// ST-FIX F23: wait until the RC left the state INITIALIZED of the previous enable
IF ( _restartReset )
THEN
  IF ( AxesGroup.Cyclic.RobToPlc.TelegramState <> TelegramState.INITIALIZED )
  THEN
    _restartReset := FALSE;
  END_IF
ELSE
CASE AxesGroup.Cyclic.RobToPlc.TelegramState  OF

         TelegramState.UNDEFINED : ;
         
         TelegramState.ERROR_161_TELEGRAM_CONTROL_MISMATCH_TELEGRAM_STATE..TelegramState.ERROR_172_TELEGRAM_NUMBER_NOT_SUPPORTED:

           // ST-FIX F79: remember the error state for the init timeout
           _initErrorState := AxesGroup.Cyclic.RobToPlc.TelegramState;

           // clear error
           AxesGroup.Cyclic.PlcToRob.Control := ControlHalfByte.ACK_ERROR;        
           AxesGroup.Cyclic.PlcToRob.Control := ControlHalfByte.RESET; // always a reset, so that on the robot side the ACR is reseted         

         TelegramState.ERROR_173_SERVER_CONNECTION_LOST:

           // Reset interface including the ACR register on server side
           AxesGroup.Cyclic.PlcToRob.Control := ControlHalfByte.RESET;        
           
         TelegramState.READY_TO_RESUME :  
         
           // Resume
           AxesGroup.Cyclic.PlcToRob.Control := ControlHalfByte.RESUME;        
         
         TelegramState.READY_FOR_INITIALIZATION: 

           // Request initialization
           AxesGroup.Cyclic.PlcToRob.Control := ControlHalfByte.INITIALIZE;
           
         TelegramState.INITIALIZED: 

           // Reset Telegram Control 
           AxesGroup.Cyclic.PlcToRob.Control := ControlHalfByte.NONE;
           
           // Check SRCI Version is compatible ? 
           IF ( AxesGroup.Cyclic.RobToPlc.SRCIVersion.MajorVersion = RobotLibraryConstants.SRCIVersion.MajorVersion )
           THEN
             // set timeout
             SetTimeout(PT := _timeoutCmd, rTimer := _timerCmd);
             // inc step counter
            _stepCmd := _stepCmd + 1; 
           ELSE
             // set error 
             ErrorID     := RobotLibraryErrorIdEnum.ERR_SRCI_MAJOR_VERSION_INCOMPATIBLE_0x80A4;
             ErrorAddTxt := CONCAT('_stepCmd = ' , DINT_TO_STRING(_stepCmd));
           END_IF

       ELSE
         // TelegrammState in error          
         SetError( ErrorID := RobotLibraryErrorIdEnum.ERR_INIT_LOST_UNKNOWN_0x80A2, Overwrite := TRUE ); // ST-FIX F65: unknown state (16#A2 is the RI error of the RC)
           // Create log entry
           CreateLogMessagePara1 ( Timestamp   := SystemTime,
                                   MessageType := MessageType.CMD,
                                   Severity    := Severity.ERROR,
                                   MessageCode := ErrorID,
                                   MessageText := 'Initialization lost: unknown telegram state {1}',
                                   Para1       := TELEGRAM_STATE_TO_STRING(AxesGroup.Cyclic.RobToPlc.TelegramState));
         ErrorAddTxt := CONCAT('_stepCmd = ' , DINT_TO_STRING(_stepCmd));
       END_CASE
END_IF

       // timeout exceeded ? 
       IF (CheckTimeout(_timerCmd) = RobotLibraryConstants.OK)
       THEN
         // Check Telegram State error ? 
         IF (( AxesGroup.Cyclic.RobToPlc.TelegramState >= TelegramState.ERROR_161_TELEGRAM_CONTROL_MISMATCH_TELEGRAM_STATE ) AND // ST-FIX F15
             ( AxesGroup.Cyclic.RobToPlc.TelegramState <= TelegramState.ERROR_173_SERVER_CONNECTION_LOST                   ))
         THEN
           ErrorID     := AxesGroup.Cyclic.RobToPlc.TelegramState;
           ErrorAddTxt := CONCAT('_stepCmd = ' , DINT_TO_STRING(_stepCmd));
         ELSIF ( _initErrorState <> TelegramState.UNDEFINED ) // ST-FIX F79: error state seen during the initialization
         THEN
           ErrorID     := _initErrorState;
           ErrorAddTxt := CONCAT('_stepCmd = ' , DINT_TO_STRING(_stepCmd));
         ELSE
           ErrorID     := RobotLibraryErrorIdEnum.ERR_TIMEOUT_CMD;
           ErrorAddTxt := CONCAT('_stepCmd = ' , DINT_TO_STRING(_stepCmd));
         END_IF
       END_IF

       
  02: IF (( NOT _readMessages.Busy  ) AND 
          ( NOT _readMessages.Error )) 
      THEN
        // start function block
       _readMessages.Enable := TRUE;
       _readMessages.ParCmd.MsgID := 0;
       _readMessages.ParCmd.MessageLevel := _parCfg.Rob.Parameter.MessageLevel;
        
        // set timeout
        SetTimeout(PT := _timeoutCmd, rTimer := _timerCmd);
        // inc step counter
       _stepCmd := _stepCmd + 1;       
      ELSE
        // check error ? 
        IF (_readMessages.Error)
        THEN
          ErrorID     := _readMessages.ErrorID;
          ErrorAddTxt := _readMessages.ErrorAddTxt;;
        END_IF  
        // timeout exceeded ? 
        IF (CheckTimeout(_timerCmd) = RobotLibraryConstants.OK)
        THEN
          ErrorID     := RobotLibraryErrorIdEnum.ERR_TIMEOUT_CMD;
          ErrorAddTxt := CONCAT('_stepCmd = ' , DINT_TO_STRING(_stepCmd));
        END_IF
      END_IF
  
  03: IF ((     _readMessages.Enabled ) AND
          ( NOT _readMessages.Error   ))
      THEN       
        // --------------------------------------------------------------- 
        // !!! ReadMessages must stay active for the Message mechanism !!!
        // --------------------------------------------------------------- 
        // ReadMessages.Enable := FALSE;  
        // set timeout
        SetTimeout(PT := _timeoutCmd, rTimer := _timerCmd);
        // inc step counter
       _stepCmd := _stepCmd + 1;
      ELSE
         // check error ? 
         IF (_readMessages.Error)
         THEN
           ErrorID     := _readMessages.ErrorID;
           ErrorAddTxt := _readMessages.ErrorAddTxt;;
         END_IF  
       
         // timeout exceeded ? 
         IF (CheckTimeout(_timerCmd) = RobotLibraryConstants.OK)
         THEN
           ErrorID     := RobotLibraryErrorIdEnum.ERR_TIMEOUT_CMD;
           ErrorAddTxt := CONCAT('_stepCmd = ' , DINT_TO_STRING(_stepCmd));
         END_IF
       END_IF       
       
       
  04: IF (( NOT _exchangeConfiguration.Busy  ) AND 
          ( NOT _exchangeConfiguration.Error ))
      THEN
        // set command parameter
       _exchangeConfiguration.ParCmd.LogLevel                           :=  LogLevel; 
       _exchangeConfiguration.ParCmd.WaitAtBlendingZone                 := _parCfg.Rob.Parameter.WaitAtBlendingZone;
       _exchangeConfiguration.ParCmd.AllowSecSeqWhileSubprogram         := _parCfg.Rob.Parameter.AllowSecSeqWhileSubprogram;
       _exchangeConfiguration.ParCmd.AllowDynamicBlending               := _parCfg.Rob.Parameter.AllowDynamicBlending;
       _exchangeConfiguration.ParCmd.DelayTime                          := _parCfg.Rob.Parameter.DelayTime;
       _exchangeConfiguration.ParCmd.WaitForNrOfCmd                     := _parCfg.Rob.Parameter.WaitForNrOfCmd;
       _exchangeConfiguration.ParCmd.LifeSignTimeOut                    :=  TIME_TO_UINT(_parCfg.Com.LifeSignTimeOut);
       _exchangeConfiguration.ParCmd.SyncDelay                          := _parCfg.Rob.Parameter.SyncDelay;
       _exchangeConfiguration.ParCmd.SyncReaction                       := _parCfg.Rob.Parameter.SyncReaction;
       _exchangeConfiguration.ParCmd.DataEnableSync                     :=  SyncModesToDataEnableSync(Value := _parCfg.Plc.Parameter.SynchronizationModes);
       _exchangeConfiguration.ParCmd.DataInSync.ToolsInSync             :=  FALSE;
       _exchangeConfiguration.ParCmd.DataInSync.FramesInSync            :=  FALSE;
       _exchangeConfiguration.ParCmd.DataInSync.LoadsInSync             :=  FALSE;
       _exchangeConfiguration.ParCmd.DataInSync.WorkAreasInSync         :=  FALSE;
       _exchangeConfiguration.ParCmd.DataInSync.SoftwareLimitsInSync    :=  FALSE;
       _exchangeConfiguration.ParCmd.DataInSync.DefaultDynamicsInSync   :=  FALSE;
       _exchangeConfiguration.ParCmd.DataInSync.ReferenceDynamicsInSync :=  FALSE;         
       
        // start function block
       _exchangeConfiguration.Enable := TRUE;
        // set timeout
        SetTimeout(PT := _timeoutCmd, rTimer := _timerCmd);
        // inc step counter
       _stepCmd := _stepCmd + 1;       
      ELSE
        // check error ? 
        IF (_exchangeConfiguration.Error)
        THEN
          ErrorID     := _exchangeConfiguration.ErrorID;
          ErrorAddTxt := _exchangeConfiguration.ErrorAddTxt;;
        END_IF  
       
        // timeout exceeded ? 
        IF (CheckTimeout(_timerCmd) = RobotLibraryConstants.OK)
        THEN
          ErrorID     := RobotLibraryErrorIdEnum.ERR_TIMEOUT_CMD;
          ErrorAddTxt := CONCAT('_stepCmd = ' , DINT_TO_STRING(_stepCmd));
        END_IF
      END_IF
  
  
  05: IF ((     _exchangeConfiguration.Enabled ) AND
          ( NOT _exchangeConfiguration.Error   ))
      THEN     
        // --------------------------------------------------------------------- 
        // !!! ExchangeConfiguration must stay active for the Sync mechanism !!!
        // --------------------------------------------------------------------- 
        // ExchangeConfiguration.Enable := FALSE;  
        // set timeout
        SetTimeout(PT := _timeoutCmd, rTimer := _timerCmd);
        // inc step counter
       _stepCmd := _stepCmd + 1;       
      ELSE
        // check error ? 
        IF (_exchangeConfiguration.Error)
        THEN
          ErrorID     := _exchangeConfiguration.ErrorID;
          ErrorAddTxt := _exchangeConfiguration.ErrorAddTxt;;
        END_IF  
       
        // timeout exceeded ? 
        IF (CheckTimeout(_timerCmd) = RobotLibraryConstants.OK)
        THEN
          ErrorID     := RobotLibraryErrorIdEnum.ERR_TIMEOUT_CMD;
          ErrorAddTxt := CONCAT('_stepCmd = ' , DINT_TO_STRING(_stepCmd));
        END_IF
      END_IF

       
  06: IF (( NOT _readRobotData.Busy  ) AND 
          ( NOT _readRobotData.Error )) 
      THEN
        // start function block
       _readRobotData.Execute := TRUE;
        // set timeout
        SetTimeout(PT := _timeoutCmd, rTimer := _timerCmd);
        // inc step counter
       _stepCmd := _stepCmd + 1;       
      ELSE
        // check error ? 
        IF (_readRobotData.Error)
        THEN
          ErrorID     := _readRobotData.ErrorID;
          ErrorAddTxt := _readRobotData.ErrorAddTxt;;
        END_IF  
        // timeout exceeded ? 
        IF (CheckTimeout(_timerCmd) = RobotLibraryConstants.OK)
        THEN
          ErrorID     := RobotLibraryErrorIdEnum.ERR_TIMEOUT_CMD;
          ErrorAddTxt := CONCAT('_stepCmd = ' , DINT_TO_STRING(_stepCmd));
        END_IF
      END_IF
    
  
  07: IF ((     _readRobotData.Done  ) AND
          ( NOT _readRobotData.Busy  ) AND
          ( NOT _readRobotData.Error ))          
      THEN       
        // set initialized flag
        Initialized := TRUE;       
        // start function block
       _readRobotData.Execute := FALSE;
        // set timeout
        SetTimeout(PT := _timeoutCmd, rTimer := _timerCmd);
        // inc step counter
       _stepCmd := _stepCmd + 1;
       ELSE
         // check error ? 
         IF (_readRobotData.Error)
         THEN
           ErrorID     := _readRobotData.ErrorID;
           ErrorAddTxt := _readRobotData.ErrorAddTxt;;
         END_IF  
       
         // timeout exceeded ? 
         IF (CheckTimeout(_timerCmd) = RobotLibraryConstants.OK)
         THEN
           ErrorID     := RobotLibraryErrorIdEnum.ERR_TIMEOUT_CMD;
           ErrorAddTxt := CONCAT('_stepCmd = ' , DINT_TO_STRING(_stepCmd));
         END_IF
       END_IF

       
  08:  // Update Initialized state
       // ST-FIX F131: Initialized stays TRUE while Synchronized (RI state "Synchronized" includes the
       // initialization); otherwise CheckParameterChanged did not run while synchronized
       Initialized := NOT Error;
       // ST-FIX F29: the next line overwrote the error check above
       // Initialized := NOT Synchronized;

       // Wait for task disable
       IF ( NOT Enable)
       THEN
         // Reset active command register
         AxesGroup.Acyclic.ActiveCommandRegister.Reset();
         // reset internal variables
         Reset(AxesGroup := AxesGroup);
         // Reset step counter
        _stepCmd := 0;         
         // finished okay
         OnExecRun := RobotLibraryConstants.OK;
       END_IF  

       
ELSE
  // invalid step
  ErrorID     := RobotLibraryErrorIdEnum.ERR_INVALID_STEP;
  ErrorAddTxt := CONCAT('_stepCmd = ' , DINT_TO_STRING(_stepCmd));
END_CASE
END_METHOD

METHOD PROTECTED ParseRecvPayload
VAR_IN_OUT
  /// Robot assignment of function
  AxesGroup   : AxesGroup;
  /// Inputs of PLC for communication from RC
  RobotInData : ARRAY[*] OF BYTE;
END_VAR
// reset all variables and payload
RecvData.Reset();
// Call RecvData FB, update payload and size 
RecvData(Payload := RobotInData, PayloadSize := ROBOT_IN_DATA_SIZE);

// check new data to receive ? 
// ST-FIX F140: also new data of the 2nd sequence
IF ( Telegram.RobToPlc.Sequence[0].Header.SEQ_ACK <> AxesGroup.State.LastACK[0] ) OR
   ( Telegram.RobToPlc.Sequence[1].Header.SEQ_ACK <> AxesGroup.State.LastACK[1] )
THEN
  // delete old telegram data 
  SysDepMemSet(pDest := ADR(Telegram.RobToPlc), Value := 0 , DataLen := SIZEOF(Telegram.RobToPlc));
END_IF


ParseRecvPayloadHeader        ( AxesGroup := AxesGroup);
ParseRecvPayloadCyclic        ( AxesGroup := AxesGroup);
ParseRecvPayloadCyclicOptional( AxesGroup := AxesGroup);
ParseRecvPayloadSequence      ( AxesGroup := AxesGroup);
ParseRecvPayloadFooter        ( AxesGroup := AxesGroup);
ParseRecvPayloadLogging       ( AxesGroup := AxesGroup);


AxesGroup.State.LastACK[0] := Telegram.RobToPlc.Sequence[0].Header.SEQ_ACK; 
AxesGroup.State.LastACK[1] := Telegram.RobToPlc.Sequence[1].Header.SEQ_ACK;
END_METHOD

METHOD PROTECTED ParseRecvPayloadCyclic
VAR_IN_OUT
  /// Robot assignment of function
  AxesGroup: AxesGroup;
END_VAR
END_METHOD

METHOD PROTECTED ParseRecvPayloadCyclicOptional
VAR_IN_OUT
  /// Robot assignment of function
  AxesGroup    : AxesGroup;
END_VAR

VAR 
  /// internal index for loops
 _idx : DINT;
END_VAR
// AxesGroup.OptionalCyclic.RobToPlc.SubProgramData {{{
IF ( AxesGroup.CyclicOptional.RobToPlc.SubProgramData.Active )
THEN
  FOR _idx := 0 TO  RobotLibraryConstants.CYCLIC_SUB_PROGRAM_DATA_MAX (* ST-FIX F179 *)
  DO
    Telegram.RobToPlc.CyclicOptional.SubProgramData.Data[_idx] := RecvData.GetByte(); 
  END_FOR
END_IF
// }}}
  
// AxesGroup.OptionalCyclic.RobToPlc.CartesianPos {{{
IF ( AxesGroup.CyclicOptional.RobToPlc.CartesianPosition.Active )
THEN
  Telegram.RobToPlc.CyclicOptional.CartesianPosition.X                    := RecvData.GetReal();
  Telegram.RobToPlc.CyclicOptional.CartesianPosition.Y                    := RecvData.GetReal();
  Telegram.RobToPlc.CyclicOptional.CartesianPosition.Z                    := RecvData.GetReal();
  Telegram.RobToPlc.CyclicOptional.CartesianPosition.Rx                   := RecvData.GetReal();
  Telegram.RobToPlc.CyclicOptional.CartesianPosition.Ry                   := RecvData.GetReal();
  Telegram.RobToPlc.CyclicOptional.CartesianPosition.Rz                   := RecvData.GetReal();
  Telegram.RobToPlc.CyclicOptional.CartesianPosition.Config               := RecvData.GetWord();
  Telegram.RobToPlc.CyclicOptional.CartesianPosition.Turns_J2_J1          := RecvData.GetByte();
  Telegram.RobToPlc.CyclicOptional.CartesianPosition.Turns_J4_J3          := RecvData.GetByte();
  Telegram.RobToPlc.CyclicOptional.CartesianPosition.Turns_J6_J5          := RecvData.GetByte();
  Telegram.RobToPlc.CyclicOptional.CartesianPosition.Turns_E1             := RecvData.GetByte();  
  Telegram.RobToPlc.CyclicOptional.CartesianPosition.E1                   := RecvData.GetReal();  
  Telegram.RobToPlc.CyclicOptional.CartesianPosition.ToolNo               := RecvData.GetUsint();
  Telegram.RobToPlc.CyclicOptional.CartesianPosition.FrameNo              := RecvData.GetUsint();
  Telegram.RobToPlc.CyclicOptional.CartesianPosition.CurrentlyUsedToolNo  := RecvData.GetUsint();
  Telegram.RobToPlc.CyclicOptional.CartesianPosition.CurrentlyUsedFrameNo := RecvData.GetUsint();
  Telegram.RobToPlc.CyclicOptional.CartesianPosition.Reserve_1            := RecvData.GetByte();
  Telegram.RobToPlc.CyclicOptional.CartesianPosition.Reserve_2            := RecvData.GetByte();  
END_IF
// }}}

// AxesGroup.OptionalCyclic.RobToPlc.JointPosition {{{
IF ( AxesGroup.CyclicOptional.RobToPlc.JointPosition.Active )
THEN
  Telegram.RobToPlc.CyclicOptional.JointPosition.J1         := RecvData.GetReal();
  Telegram.RobToPlc.CyclicOptional.JointPosition.J2         := RecvData.GetReal();
  Telegram.RobToPlc.CyclicOptional.JointPosition.J3         := RecvData.GetReal();
  Telegram.RobToPlc.CyclicOptional.JointPosition.J4         := RecvData.GetReal();
  Telegram.RobToPlc.CyclicOptional.JointPosition.J5         := RecvData.GetReal();
  Telegram.RobToPlc.CyclicOptional.JointPosition.J6         := RecvData.GetReal();
  Telegram.RobToPlc.CyclicOptional.JointPosition.E1         := RecvData.GetReal();
  Telegram.RobToPlc.CyclicOptional.JointPosition.E1_Reserve := RecvData.GetWord();
END_IF  
// }}}

// AxesGroup.OptionalCyclic.RobToPlc.CartesianForce {{{
IF ( AxesGroup.CyclicOptional.RobToPlc.Force.Active )
THEN
  Telegram.RobToPlc.CyclicOptional.Force.X  := RecvData.GetReal();
  Telegram.RobToPlc.CyclicOptional.Force.Y  := RecvData.GetReal();
  Telegram.RobToPlc.CyclicOptional.Force.Z  := RecvData.GetReal();
  Telegram.RobToPlc.CyclicOptional.Force.Rx := RecvData.GetReal();
  Telegram.RobToPlc.CyclicOptional.Force.Ry := RecvData.GetReal();
  Telegram.RobToPlc.CyclicOptional.Force.Rz := RecvData.GetReal();
END_IF  
// }}}    
  
// AxesGroup.OptionalCyclic.RobToPlc.Current {{{
IF ( AxesGroup.CyclicOptional.RobToPlc.Current.Active )
THEN
  Telegram.RobToPlc.CyclicOptional.Current.J1  := RecvData.GetReal();
  Telegram.RobToPlc.CyclicOptional.Current.J2  := RecvData.GetReal();
  Telegram.RobToPlc.CyclicOptional.Current.J3  := RecvData.GetReal();
  Telegram.RobToPlc.CyclicOptional.Current.J4  := RecvData.GetReal();
  Telegram.RobToPlc.CyclicOptional.Current.J5  := RecvData.GetReal();
  Telegram.RobToPlc.CyclicOptional.Current.J6  := RecvData.GetReal();
END_IF    
  
// AxesGroup.OptionalCyclic.RobToPlc.CartesianPosExt {{{
IF ( AxesGroup.CyclicOptional.RobToPlc.CartesianPositionExt.Active )
THEN
  Telegram.RobToPlc.CyclicOptional.CartesianPositionExt.E2 := RecvData.GetReal();
  Telegram.RobToPlc.CyclicOptional.CartesianPositionExt.E3 := RecvData.GetReal();
  Telegram.RobToPlc.CyclicOptional.CartesianPositionExt.E4 := RecvData.GetReal();
  Telegram.RobToPlc.CyclicOptional.CartesianPositionExt.E5 := RecvData.GetReal();
  Telegram.RobToPlc.CyclicOptional.CartesianPositionExt.E6 := RecvData.GetReal();
END_IF  
// }}}       
  
// AxesGroup.OptionalCyclic.RobToPlc.JointPosition {{{
IF ( AxesGroup.CyclicOptional.RobToPlc.JointPositionExt.Active )
THEN
  Telegram.RobToPlc.CyclicOptional.JointPositionExt.E2 := RecvData.GetReal();
  Telegram.RobToPlc.CyclicOptional.JointPositionExt.E3 := RecvData.GetReal();
  Telegram.RobToPlc.CyclicOptional.JointPositionExt.E4 := RecvData.GetReal();
  Telegram.RobToPlc.CyclicOptional.JointPositionExt.E5 := RecvData.GetReal();
  Telegram.RobToPlc.CyclicOptional.JointPositionExt.E6 := RecvData.GetReal();  
END_IF  
// }}}    
      
// AxesGroup.OptionalCyclic.RobToPlc.CartesianForceExt {{{
IF ( AxesGroup.CyclicOptional.RobToPlc.ForceExt.Active )
THEN
  Telegram.RobToPlc.CyclicOptional.ForceExt.E1  := RecvData.GetReal();
  Telegram.RobToPlc.CyclicOptional.ForceExt.E2  := RecvData.GetReal();
  Telegram.RobToPlc.CyclicOptional.ForceExt.E3  := RecvData.GetReal();
  Telegram.RobToPlc.CyclicOptional.ForceExt.E4  := RecvData.GetReal();
  Telegram.RobToPlc.CyclicOptional.ForceExt.E5  := RecvData.GetReal();
  Telegram.RobToPlc.CyclicOptional.ForceExt.E6  := RecvData.GetReal();
END_IF
// }}}    
  
// AxesGroup.OptionalCyclic.RobToPlc.CurrentExt {{{
IF ( AxesGroup.CyclicOptional.RobToPlc.CurrentExt.Active )
THEN
  Telegram.RobToPlc.CyclicOptional.CurrentExt.E1  := RecvData.GetReal();
  Telegram.RobToPlc.CyclicOptional.CurrentExt.E2  := RecvData.GetReal();
  Telegram.RobToPlc.CyclicOptional.CurrentExt.E3  := RecvData.GetReal();
  Telegram.RobToPlc.CyclicOptional.CurrentExt.E4  := RecvData.GetReal();
  Telegram.RobToPlc.CyclicOptional.CurrentExt.E5  := RecvData.GetReal();
  Telegram.RobToPlc.CyclicOptional.CurrentExt.E6  := RecvData.GetReal();
END_IF
// }}}
END_METHOD

METHOD PRIVATE ParseRecvPayloadFooter
VAR_IN_OUT
  /// Robot assignment of function
  AxesGroup : AxesGroup;
END_VAR
Telegram.RobToPlc.Footer.LifeSign := RecvData.GetLifeSignFooter();
END_METHOD

METHOD PROTECTED ParseRecvPayloadHeader
VAR_IN_OUT
  /// Robot assignment of function
  AxesGroup    : AxesGroup;
END_VAR
// Version
Telegram.RobToPlc.Header.SRCIVersion := ByteToVersion(RecvData.GetByte());
// Connection alive signal
Telegram.RobToPlc.Header.LifeSign    := RecvData.GetHalfeByte2(IncPayloadPtr := TRUE);
// Reserved byte
Telegram.RobToPlc.Header.Reserved       := RecvData.GetByte();
// Initialization and Telegram control state
Telegram.RobToPlc.Header.TelegramState  := RecvData.GetUsint();
// Combination of various RA related states.
Telegram.RobToPlc.Header.StatusRobotArm := RecvData.GetDword();
// Actual override in percentage encoding 
Telegram.RobToPlc.Header.Override       := RecvData.GetUint();
END_METHOD

METHOD PRIVATE ParseRecvPayloadLogging
VAR_IN_OUT
  /// Robot assignment of function
  AxesGroup    : AxesGroup;
END_VAR

VAR
  /// internal sequence index for loops
  _seqIdx : DINT;
  /// internal fragment index for loops
  _fragIdx : DINT;
END_VAR
RETURN;
FOR _seqIdx := 0 TO AxesGroup.State.SequenceCountRecv
DO
  // check new data to receive ? 
  IF ( Telegram.RobToPlc.Sequence[_seqIdx].Header.SEQ_ACK <> AxesGroup.State.LastACK[_seqIdx]) 
  THEN
    // Check sequence payload > 0 ?    
    IF (Telegram.RobToPlc.Sequence[_seqIdx].Header.PayloadLength > 0)
    THEN
      // Create log entry
      CreateLogMessagePara4 ( Timestamp   := SystemTime,
                              MessageType := MessageType.CMD,
                              Severity    := Severity.DEBUG,
                              MessageCode := 0,
                              MessageText := 'RecvData: ACK = {1}, received Sequence [{2}] with PayloadLength = {3}, Lifesign = {4}',
                              Para1       :=  UINT_TO_STRING(Telegram.RobToPlc.Sequence[_seqIdx].Header.SEQ_ACK),
                              Para2       :=  DINT_TO_STRING(_seqIdx),
                              Para3       :=  UINT_TO_STRING(Telegram.RobToPlc.Sequence[_seqIdx].Header.PayloadLength),
                              Para4       :=  BYTE_TO_STRING(Telegram.RobToPlc.Header.LifeSign));
  
      FOR _fragIdx := 0 TO AxesGroup.State.FragmentCountRecv[_seqIdx] 
      DO
        // Check fragment payload > 0 ?    
        IF (Telegram.RobToPlc.Sequence[_seqIdx].Fragment[_fragIdx].Header.PayloadLength > 0)
        THEN
          // Create log entry
          CreateLogMessagePara5 ( Timestamp   := SystemTime,
                                  MessageType := MessageType.CMD,
                                  Severity    := Severity.DEBUG,
                                  MessageCode := 0,
                                  MessageText := 'RecvData: received Fragment [{1}] with PayloadLength = {2}, CmdID <{3}> , CmdState: {4}, Fragment-Action Bits: {5}',
                                  Para1       :=  DINT_TO_STRING(_fragIdx),
                                  Para2       :=  UINT_TO_STRING              (Telegram.RobToPlc.Sequence[_seqIdx].Fragment[_fragIdx].Header.PayloadLength),
                                  Para3       :=  DINT_TO_STRING              (Telegram.RobToPlc.Sequence[_seqIdx].Fragment[_fragIdx].Header.CmdID),
                                  Para4       :=  CMD_MESSAGE_STATE_TO_STRING (Telegram.RobToPlc.Sequence[_seqIdx].Fragment[_fragIdx].Command.Header.State),
                                  Para5       :=    FRAGMENT_ACTION_TO_STRING (Telegram.RobToPlc.Sequence[_seqIdx].Fragment[_fragIdx].Header.FragmentAction));
        END_IF
      END_FOR    
    END_IF
  END_IF
END_FOR
END_METHOD

METHOD PRIVATE ParseRecvPayloadSequence
VAR_IN_OUT
  /// Robot assignment of function
  AxesGroup        : AxesGroup;
END_VAR

VAR
  /// internal index
 _idx              : DINT;
  /// index for sequence
 _seqIdx           : DINT;
  /// index for fragment
 _fragIdx          : DINT; 
  /// current payload pointer for current fragment
 _payLoadPtr       : DINT;
  /// Amount of sequences
 _seqCount         : DINT;
  /// current payload pointer of the current sequence
 _seqPayloadPtr    : UINT; 
  /// ST-FIX F63: start of the payload of each sequence (behind its sequence header)
 _rcvStart         : ARRAY[0..1] OF DINT;
  /// ST-FIX F63: sequence that is processed first (lower Ack)
 _rcvFirst         : DINT;
  /// ST-FIX F63: loop counter over the sequences in Ack order
 _rcvOrderIdx      : DINT;
  /// ST-FIX F63: distance of the two Ack numbers
 _rcvDiff          : DINT;
END_VAR
// Check 2nd sequence active ? 
IF ( _parCfg.Com.TwoSequences )
THEN
 _seqCount := _seqCount + 1;
END_IF

// ST-FIX F63: read the headers of all sequences, each from its own address (Fig. 5-205)
FOR _seqIdx := 0 TO _seqCount
DO
  IF ( _seqIdx = PRIMARY_SEQUENCE )
  THEN
    RecvData.PayloadPtr := CalculateSequencePayloadStartAdr(AxesGroup := AxesGroup, 
                                                            Direction := ComDirection.ROB_TO_PLC,
                                                            Sequence  := SequenceFlag.PRIMARY_SEQUENCE);
  ELSE
    RecvData.PayloadPtr := CalculateSequencePayloadStartAdr(AxesGroup := AxesGroup, 
                                                            Direction := ComDirection.ROB_TO_PLC,
                                                            Sequence  := SequenceFlag.SECONDARY_SEQUENCE);
  END_IF

  // parse sequence header
  Telegram.RobToPlc.Sequence[_seqIdx].Header.SEQ_ACK       := RecvData.GetUint();
  Telegram.RobToPlc.Sequence[_seqIdx].Header.PayloadLength := RecvData.GetUint();
 _rcvStart[_seqIdx] := RecvData.PayloadPtr;
END_FOR

// ST-FIX F63: the sequence with the lower Ack first (Fig. 5-207/5-208), numbers wrap 254 -> 1
_rcvFirst := 0;
IF ( _seqCount = 1 )
THEN
 _rcvDiff := UINT_TO_DINT(Telegram.RobToPlc.Sequence[0].Header.SEQ_ACK)
           - UINT_TO_DINT(Telegram.RobToPlc.Sequence[1].Header.SEQ_ACK);
  IF ( _rcvDiff < 0 ) THEN _rcvDiff := _rcvDiff + 254; END_IF
  IF (( _rcvDiff > 0 ) AND ( _rcvDiff < 127 )) THEN _rcvFirst := 1; END_IF
END_IF

FOR _rcvOrderIdx := 0 TO _seqCount
DO
  IF ( _rcvOrderIdx = 0 ) THEN _seqIdx := _rcvFirst; ELSE _seqIdx := 1 - _rcvFirst; END_IF

  // ST-FIX F5: every sequence starts with fragment 0
  _fragIdx       := 0;
  _seqPayloadPtr := 0;
  RecvData.PayloadPtr := _rcvStart[_seqIdx];
  
  // check new data available ? 
  // ST-FIX F63: only the Ack of the Seq that was sent (Seq = Ack) carries the response of it;
  // with two sequences the RC may send Ack 0 in the sequence it does not process
  IF (( Telegram.RobToPlc.Sequence[_seqIdx].Header.SEQ_ACK <> AxesGroup.State.LastACK[_seqIdx]    ) AND
      ( Telegram.RobToPlc.Sequence[_seqIdx].Header.SEQ_ACK  = AxesGroup.State.CurrentSEQ[_seqIdx] ))
  THEN
    // Check sequence payload available ? 
    IF (Telegram.RobToPlc.Sequence[_seqIdx].Header.PayloadLength > 0)
    THEN
      // Check sequence payload length is valid ? 
      IF ( Telegram.RobToPlc.Sequence[_seqIdx].Header.PayloadLength > _parCfg.Com.TelegramLengthRobToPlc )
      THEN 
        // Create log entry for payload not valid 
        CreateLogMessagePara2 ( Timestamp   := SystemTime,
                                MessageType := MessageType.CMD,
                                Severity    := Severity.DEBUG,
                                MessageCode := 0,
                                MessageText := 'Invalid sequence payload length, Sequence = {1}, PayloadLength = {2} ',
                                Para1       :=  DINT_TO_STRING(_seqIdx),
                                Para2       :=  UINT_TO_STRING(Telegram.RobToPlc.Sequence[_seqIdx].Header.PayloadLength));
                                RETURN;
      ELSE
        // Create log entry
        CreateLogMessagePara4 ( Timestamp   := SystemTime,
                                MessageType := MessageType.CMD,
                                Severity    := Severity.DEBUG,
                                MessageCode := 0,
                                MessageText := 'RecvData: ACK = {1}, received Sequence [{2}] with PayloadLength = {3}, Lifesign = {4}',
                                Para1       :=  UINT_TO_STRING(Telegram.RobToPlc.Sequence[_seqIdx].Header.SEQ_ACK),
                                Para2       :=  DINT_TO_STRING(_seqIdx),
                                Para3       :=  UINT_TO_STRING(Telegram.RobToPlc.Sequence[_seqIdx].Header.PayloadLength),
                                Para4       :=  BYTE_TO_STRING(Telegram.RobToPlc.Header.LifeSign));
      END_IF
    
      // processing sequence payload                                  
      WHILE ( _seqPayloadPtr < Telegram.RobToPlc.Sequence[_seqIdx].Header.PayloadLength )
      DO                        
        // parse header
        Telegram.RobToPlc.Sequence[_seqIdx].Fragment[_fragIdx].Header.CmdID          := RecvData.GetUint();
        Telegram.RobToPlc.Sequence[_seqIdx].Fragment[_fragIdx].Header.Reserve        := RecvData.GetByte();
        Telegram.RobToPlc.Sequence[_seqIdx].Fragment[_fragIdx].Header.FragmentAction := RecvData.GetByte();
        Telegram.RobToPlc.Sequence[_seqIdx].Fragment[_fragIdx].Header.PayloadPointer := RecvData.GetUint();
        Telegram.RobToPlc.Sequence[_seqIdx].Fragment[_fragIdx].Header.PayloadLength  := RecvData.GetUint();
       
        // add header size to payload pointer 
       _seqPayloadPtr := _seqPayloadPtr + SIZEOF(Telegram.RobToPlc.Sequence[_seqIdx].Fragment[_fragIdx].Header);
        
        // Check fragment payload available ? 
        IF (Telegram.RobToPlc.Sequence[_seqIdx].Fragment[_fragIdx].Header.PayloadLength > 0)
        THEN
          // Check fragment payload length is valid ? 
          IF ( Telegram.RobToPlc.Sequence[_seqIdx].Fragment[_fragIdx].Header.PayloadLength > _parCfg.Com.TelegramLengthRobToPlc )
          THEN 
            // Create log entry for payload not valid 
            CreateLogMessagePara2 ( Timestamp   := SystemTime,
                                    MessageType := MessageType.CMD,
                                    Severity    := Severity.DEBUG,
                                    MessageCode := 0,
                                    MessageText := 'Invalid fragment payload length, Sequence = {1}, PayloadLength = {2} ',
                                    Para1       :=  DINT_TO_STRING(_seqIdx),
                                    Para2       :=  UINT_TO_STRING(Telegram.RobToPlc.Sequence[_seqIdx].Fragment[_fragIdx].Header.PayloadLength));
                                    RETURN;
          END_IF
        
          // Fill Response payload
          FOR _idx := 0 TO Telegram.RobToPlc.Sequence[_seqIdx].Fragment[_fragIdx].Header.PayloadLength -1
          DO
            // calculate payload pointer
           _payLoadPtr := Telegram.RobToPlc.Sequence[_seqIdx].Fragment[_fragIdx].Header.PayloadPointer + _idx;
          
            IF (( _payLoadPtr >= 0                                          ) AND
                ( _payLoadPtr <= RobotLibraryParameter.RESPONSE_PAYLOAD_MAX ))
            THEN  
              Telegram.RobToPlc.Sequence[_seqIdx].Fragment[_fragIdx].Command.Payload[_payLoadPtr] := RecvData.GetByte();
              // inc payload pointer
             _seqPayloadPtr := _seqPayloadPtr + SIZEOF(BYTE);
            ELSE
              // Create log entry for payload pointer not valid 
              CreateLogMessagePara3 ( Timestamp   := SystemTime,
                                      MessageType := MessageType.CMD,
                                      Severity    := Severity.DEBUG,
                                      MessageCode := 0,
                                      MessageText := 'Invalid fragment payload pointer, Sequence = {1}, Fragment = {2}, PayloadPointer = {3} ',
                                      Para1       :=  DINT_TO_STRING(_seqIdx),
                                      Para2       :=  DINT_TO_STRING(_fragIdx),
                                      Para3       :=  DINT_TO_STRING(_payLoadPtr));
                                      RETURN;
					  END_IF
           
          END_FOR
          
          // Add Response to ACR
          AxesGroup.Acyclic.ActiveCommandRegister.AddRsp(Telegram.RobToPlc.Sequence[_seqIdx].Fragment[_fragIdx]);
        
          // Only for debugging - header is part of the payload itself
          Telegram.RobToPlc.Sequence[_seqIdx].Fragment[_fragIdx].Command.Header.State                 :=      GetHalfeByteLo( Value :=  Telegram.RobToPlc.Sequence[_seqIdx].Fragment[_fragIdx].Command.Payload[0]);
          Telegram.RobToPlc.Sequence[_seqIdx].Fragment[_fragIdx].Command.Header.ParSeq                :=      GetHalfeByteHi( Value :=  Telegram.RobToPlc.Sequence[_seqIdx].Fragment[_fragIdx].Command.Payload[0]);
          Telegram.RobToPlc.Sequence[_seqIdx].Fragment[_fragIdx].Command.Header.AlarmMessageSeverity  :=        BYTE_TO_SINT(           Telegram.RobToPlc.Sequence[_seqIdx].Fragment[_fragIdx].Command.Payload[1]);
          Telegram.RobToPlc.Sequence[_seqIdx].Fragment[_fragIdx].Command.Header.AlarmMessageCode      :=  CombineBytesToUint( HiByte := Telegram.RobToPlc.Sequence[_seqIdx].Fragment[_fragIdx].Command.Payload[2],
                                                                                                                              LoByte := Telegram.RobToPlc.Sequence[_seqIdx].Fragment[_fragIdx].Command.Payload[3]);
          // Create log entry
          CreateLogMessagePara5 ( Timestamp   := SystemTime,
                                  MessageType := MessageType.CMD,
                                  Severity    := Severity.DEBUG,
                                  MessageCode := 0,
                                  MessageText := 'RecvData: received Fragment [{1}] with PayloadLength = {2}, CmdID <{3}> , CmdState: {4}, Fragment-Action Bits: {5}',
                                  Para1       :=  DINT_TO_STRING(_seqIdx),
                                  Para2       :=  UINT_TO_STRING              (Telegram.RobToPlc.Sequence[_seqIdx].Fragment[_fragIdx].Header.PayloadLength),
                                  Para3       :=  DINT_TO_STRING              (Telegram.RobToPlc.Sequence[_seqIdx].Fragment[_fragIdx].Header.CmdID),
                                  Para4       :=  CMD_MESSAGE_STATE_TO_STRING (Telegram.RobToPlc.Sequence[_seqIdx].Fragment[_fragIdx].Command.Header.State),
                                  Para5       :=    FRAGMENT_ACTION_TO_STRING (Telegram.RobToPlc.Sequence[_seqIdx].Fragment[_fragIdx].Header.FragmentAction));
        END_IF
        
        // Check still payload left ? -> goto next fragment  
        IF ( _seqPayloadPtr < Telegram.RobToPlc.Sequence[_seqIdx].Header.PayloadLength )
        THEN
         _fragIdx := _fragIdx + 1;        
        END_IF
        
        // Check fragment index limit reached ? 
        IF ( _fragIdx > RobotLibraryParameter.FRAGMENT_MAX ) 
        THEN 
          // Create log entry
          CreateLogMessagePara1 ( Timestamp   := SystemTime,
                                  MessageType := MessageType.CMD,
                                  Severity    := Severity.ERROR, // ST-FIX F52: responses are lost
                                  MessageCode := 0,
                                  MessageText := 'Fragment index out of range, _fragIdx = {1} ',
                                  Para1       :=  DINT_TO_STRING(_fragIdx));
                                  RETURN;
        END_IF        
      END_WHILE    
    END_IF
  END_IF    
END_FOR
END_METHOD

METHOD Reset
VAR_IN_OUT
  /// Robot assignment of function
  AxesGroup : AxesGroup;  
END_VAR
// reset flags
Busy              := FALSE;
Initialized       := FALSE;
Synchronized      := FALSE;
Error             := FALSE;
ErrorID           := 0;
ErrorAddTxt       := '';
WarningID         := 0;
InfoID            := 0;  

// Reset internal functon blocks
_exchangeConfiguration      .Enable  := FALSE;
_readRobotData              .Execute := FALSE;
_readMessages               .Enable  := FALSE;  
_readToolData               .Execute := FALSE;  
_readFrameData              .Execute := FALSE;  
_readLoadData               .Execute := FALSE;  
_readWorkArea               .Execute := FALSE;  
_readRobotSWLimits          .Execute := FALSE;  
_readRobotDefaultDynamics   .Execute := FALSE;  
_readRobotReferenceDynamics .Execute := FALSE;  
_writeToolData              .Execute := FALSE;   
_writeFrameData             .Execute := FALSE;   
_writeLoadData              .Execute := FALSE;   
_writeWorkArea              .Execute := FALSE;   
_writeRobotSWLimits         .Execute := FALSE;   
_writeRobotDefaultDynamics  .Execute := FALSE;   
_writeRobotReferenceDynamics.Execute := FALSE;   

// Set Client error to force server error
AxesGroup.Cyclic.PlcToRob.Control := ControlHalfByte.NONE;

// Reset synchronisation state variables
AxesGroup.State.SyncStatePlc.InSync.Frame             := FALSE;
AxesGroup.State.SyncStatePlc.InSync.Tool              := FALSE;
AxesGroup.State.SyncStatePlc.InSync.Load              := FALSE;
AxesGroup.State.SyncStatePlc.InSync.WorkArea          := FALSE;
AxesGroup.State.SyncStatePlc.InSync.SwLimits          := FALSE;
AxesGroup.State.SyncStatePlc.InSync.DefaultDynamics   := FALSE;
AxesGroup.State.SyncStatePlc.InSync.ReferenceDynamics := FALSE;

AxesGroup.State.SyncStatePlc.UnSyncNo.Frame    := 0;
AxesGroup.State.SyncStatePlc.UnSyncNo.Tool     := 0;
AxesGroup.State.SyncStatePlc.UnSyncNo.Load     := 0;
AxesGroup.State.SyncStatePlc.UnSyncNo.WorkArea := 0;

AxesGroup.State.SyncStateRc .InSync.Frame             := FALSE;
AxesGroup.State.SyncStateRc .InSync.Tool              := FALSE;
AxesGroup.State.SyncStateRc .InSync.Load              := FALSE;
AxesGroup.State.SyncStateRc .InSync.WorkArea          := FALSE;
AxesGroup.State.SyncStateRc .InSync.SwLimits          := FALSE;
AxesGroup.State.SyncStateRc .InSync.DefaultDynamics   := FALSE;
AxesGroup.State.SyncStateRc .InSync.ReferenceDynamics := FALSE;

AxesGroup.State.SyncStateRc .UnSyncNo.Frame    := 0;
AxesGroup.State.SyncStateRc .UnSyncNo.Tool     := 0;
AxesGroup.State.SyncStateRc .UnSyncNo.Load     := 0;
AxesGroup.State.SyncStateRc .UnSyncNo.WorkArea := 0;

// Reset active command register
AxesGroup.Acyclic.ActiveCommandRegister.Reset();
      
// reset step counters
_stepCmd                   := 0;
_stepSyncFrameData         := 0;
_stepSyncLoadData          := 0;
_stepSyncDefaultDynamics   := 0;
_stepSyncReferenceDynamics := 0;
_stepSyncSWLimits          := 0;
_stepSyncToolData          := 0;
_stepSyncWorkArea          := 0;
END_METHOD

METHOD PUBLIC SetError
VAR_INPUT
  /// ErrorID reported by RC for error identification according to Table 7-1
  ErrorID   : WORD;
  /// TRUE = overwrite an existing error 
  Overwrite : BOOL;
END_VAR
IF ( NOT HasError ) OR ( Overwrite )
THEN
  THIS^.ErrorID := ErrorID;
END_IF
END_METHOD

METHOD PUBLIC SetInfo
VAR_INPUT
  /// InfoID for info identification reported during execution of command according to Table 7-5
  InfoID    : WORD;
  /// TRUE = overwrite an existing info 
  Overwrite : BOOL;
END_VAR
IF ( NOT HasInfo ) OR ( Overwrite )
THEN
  THIS^.InfoID := InfoID;
END_IF
END_METHOD

METHOD PUBLIC SetWarning
VAR_INPUT
  /// WarningID for warning identification reported during execution of command according to Table 7-3
  WarningID : WORD;
  /// TRUE = overwrite an existing warning 
  Overwrite : BOOL;
END_VAR
IF ( NOT HasWarning ) OR ( Overwrite )
THEN
  THIS^.WarningID := WarningID;
END_IF
END_METHOD

/// ST-FIX F130: TRUE when the synchronization modes of a data set are defined
/// (during the start-up NO_SYNCHRONIZATION .. SERVER_TO_CLIENT, after the start-up also AUTOMATIC)
METHOD PRIVATE SyncModesValid : BOOL
VAR_INPUT
  /// Synchronization mode during the start-up
  During : SyncMode;
  /// Synchronization mode after the start-up
  After  : SyncMode;
END_VAR
SyncModesValid := ( During >= SyncMode.NO_SYNCHRONIZATION ) AND
                  ( During <  SyncMode.AUTOMATIC          ) AND
                  ( After  >= SyncMode.NO_SYNCHRONIZATION ) AND
                  ( After  <= SyncMode.AUTOMATIC          );
END_METHOD

END_FUNCTION_BLOCK

// Library/POUs/Read/MC_ReadToolData/MC_ReadToolDataFB

            
              /// Read content of selected tool number
FUNCTION_BLOCK MC_ReadToolDataFB EXTENDS RobotLibraryBaseExecuteFB
// ------------------------------------------------------------------------- 
//  SRCI Robot Library                                                
// ------------------------------------------------------------------------- 
//                                                                           
//  Object:      ReadToolDataFB                                       
//  Author:      Thorsten Brach                                                
//  Date:        2024-06-01
//
//  Description:                                              
//   
//                                                                           
//  Copyright: 
//    (C) 2024 Thorsten Brach. All rights reserved                                                                                                                                            
//             Licensed under the MIT License.
//                                                                           
//  Disclaimer:                                                                           
//    This project is provided without any guarantee and can be used for   
//    private and commercial purposes. Any use is at the user’s 
//    own risk and responsibility.
//
// -------------------------------------------------------------------------
VAR_INPUT
  /// command parameter 
  ParCmd          : ReadToolDataParCmd;
END_VAR
VAR_OUTPUT
  /// Command is transferred and confirmed by the RC
  CommandBuffered : BOOL;
  /// command outputs
  OutCmd          : ReadToolDataOutCmd;       
END_VAR

VAR
  /// internal copy of command parameter 
 _parCmd          : ReadToolDataParCmd;
  /// command data to send
 _command         : ReadToolDataSendData;
  /// response data received
 _response        : ReadToolDataRecvData;      
END_VAR

            
          
VAR_INPUT
  UpdateSystemData : BOOL := TRUE; // ST-FIX F16: FALSE for the internal instances of MC_RobotTaskFB (synchronisation)
END_VAR

SUPER^(AxesGroup := AxesGroup);

METHOD INTERNAL CheckAddParameter : BOOL
VAR_INPUT
  /// Payload pointer
  PayloadPtr : UDINT;
END_VAR
VAR
  /// Payload as byte array
  Payload    : ARRAY [1..SIZEOF(_command)] OF BYTE;
  /// Null Byte array 
  Null       : ARRAY [1..SIZEOF(_command)] OF BYTE;
  /// Data length to compare
  DataLen    : UDINT;
END_VAR
// Payload pointer must be decreased by one byte, because ADR(Payload) is already one byte !
PayloadPtr := LIMIT (0, PayloadPtr - 1, SIZEOF(Payload) -1);
// Convert command struct to payload array
SysDepMemCpy( pDest := ADR(Payload), pSrc := ADR(_command), DataLen := SIZEOF(_command));
// Calculate the data length to compare - at least one byte must be compared !
DataLen := LIMIT(1, SIZEOF(Payload) - PayloadPtr, SIZEOF(Payload)); 
// Compare Payload-Array with Null-Byte-Array
CheckAddParameter := SysDepMemCmp( pData1 := ADR(Payload) + PayloadPtr , pData2 := ADR(Null), DataLen := DataLen) <>  RobotLibraryConstants.OK ;
END_METHOD

METHOD PROTECTED CheckFunctionSupported : BOOL
VAR_IN_OUT
  /// Robot assignment of function
  AxesGroup : AxesGroup; 
END_VAR
CheckFunctionSupported := AxesGroup.State.RobotData.RCSupportedFunctions.ReadToolData;

IF ( NOT CheckFunctionSupported )
THEN
  // call base implementation for set error and create log entry
  SUPER^.CheckFunctionSupported(AxesGroup := AxesGroup);
END_IF
END_METHOD

METHOD PROTECTED CheckParameterChanged : BOOL
VAR_IN_OUT
  /// Robot assignment of function
  AxesGroup    : AxesGroup; 
END_VAR
// Check ParCmd Size is > 0, because MemCmp does not work correctly with size = 0
IF (SIZEOF(ParCmd) = 0) OR (_stepCmd = 0)
THEN 
  RETURN;
END_IF

// compare memory 
_parameterChanged := ( SysDepMemCmp(pData1 := ADR(ParCmd), pData2 := ADR(_parCmd), DataLen := SIZEOF(ParCmd)) <> RobotLibraryConstants.OK );

// check parameter valid ?
_parameterValid   := CheckParameterValid( AxesGroup := AxesGroup );

IF ((  _parameterChanged        )  AND 
    (  _parameterValid          )) OR
    (  _parameterUpdateInternal )  
THEN  
  // Create log entry for parameter changed event
  CreateLogMessagePara1 ( Timestamp   := AxesGroup.State.SystemTime,
                          MessageType := MessageType.CMD,
                          Severity    := Severity.DEBUG,
                          MessageCode := 0,
                          MessageText := 'NotifyParameterChanged Event {1}',
                          Para1       :=  '' );

  // reset internal flag for send parameter update
 _parameterUpdateInternal := FALSE;
  // update internal copy of parameters 
 _parCmd := ParCmd;
  // inc parameter sequence
 _command.ParSeq := _command.ParSeq + 1;
  // update command data  
  CommandData := CreateCommandPayload(AxesGroup := AxesGroup); // ( Access via reference to rCommandFB in ACR )
  // notify active command register 
  AxesGroup.Acyclic.ActiveCommandRegister.NotifyParameterChanged := _uniqueID;
END_IF
END_METHOD

METHOD PROTECTED CheckParameterValid : BOOL
VAR_IN_OUT
  /// Robot assignment of function
  AxesGroup : AxesGroup; 
END_VAR
VAR
  /// internal index for loops
 _idx : DINT;
END_VAR
CheckParameterValid := TRUE;

// Check ParCmd.ToolNo valid ? 
IF (( ParCmd.ToolNo <  -1                                                ) OR  
    ( ParCmd.ToolNo > 254                                                ) OR
    ( ParCmd.ToolNo > AxesGroup.State.ConfigurationData.HighestToolIndex ) OR
    ( ParCmd.ToolNo > AxesGroup.State.UnifiedToolIndex                   ))
THEN
  // Parameter not valid
  CheckParameterValid := FALSE;
  
  // Check ToolNo available on RC ? 
  IF (( ParCmd.ToolNo > AxesGroup.State.ConfigurationData.HighestToolIndex ) AND ( ParCmd.ToolNo <= 254 )) // ST-FIX F98: outside -1..254 is a range error
  THEN
    SetError( ErrorID := RobotLibraryErrorIdEnum.ERR_TOOLNO_UNAVAILABLE, Overwrite := TRUE );
  ELSE
    SetError( ErrorID := RobotLibraryErrorIdEnum.ERR_TOOLNO_RANGE, Overwrite := TRUE );
	END_IF  
  
  // Create log entry
  CreateLogMessagePara1 ( Timestamp   := AxesGroup.State.SystemTime,
                          MessageType := MessageType.CMD,
                          Severity    := Severity.ERROR,
                          MessageCode := ErrorID,
                          MessageText := 'Invalid Parameter ParCmd.ToolNo = {1}',
                          Para1       :=  INT_TO_STRING(ParCmd.ToolNo));
  RETURN;                          
END_IF
END_METHOD

METHOD INTERNAL CreateCommandPayload : RobotLibraryCommandDataFB
VAR_IN_OUT
  /// Robot assignment of function
  AxesGroup : AxesGroup; 
END_VAR
VAR
  /// Parameter count
 _parameterCnt : DINT;
END_VAR
// Table 6-189: Sent CMD payload (PLC to RC) of "ReadToolData"
// --------------------------
// Header
// --------------------------
// Byte 00 : UINT  - Type HB     
// Byte 01 :       - Type LB    
// Byte 02 : USINT - Reserve | ExecutionMode
// Byte 03 : USINT - ParSeq  | Priority
// --------------------------
// Datablock
// --------------------------
// Byte 04 : USINT - ToolNo;
// --------------------------
// set command parameter 
_command.CmdTyp   :=  CmdType.ReadToolData;
_command.ExecMode :=  ExecMode;
_command.ParSeq   := _command.ParSeq;
_command.Priority :=  Priority;
_command.ToolNo   := INT_TO_USINT(_parCmd.ToolNo);

IF (_parCmd.ToolNo = -1)
THEN
  _command.ToolNo := 255;
END_IF

// copy command data to header
_cmdHeader := _command;
// call base implementation to copy header to payload buffer
CreateCommandPayload := SUPER^.CreateCommandPayload(AxesGroup := AxesGroup);


// Check parameter must be added ? 
IF ( CheckAddParameter(CreateCommandPayload.PayloadPtr))
THEN
  // add command.ToolNo
  CreateCommandPayload.AddUsint(_command.ToolNo);
  // inc parameter counter
 _parameterCnt := _parameterCnt + 1;  
END_IF


// Create logging
CreateCommandPayloadLog(AxesGroup := AxesGroup, ParameterCnt := _parameterCnt);
END_METHOD

METHOD INTERNAL CreateCommandPayloadLog
VAR_IN_OUT
  /// Robot assignment of function
  AxesGroup : AxesGroup; 
END_VAR
VAR_INPUT
  /// Parameter count
  ParameterCnt : DINT;
END_VAR
// Create log entry for Parameter start
CreateLogMessagePara1 ( Timestamp   := AxesGroup.State.SystemTime,
                        MessageType := MessageType.CMD,
                        Severity    := Severity.DEBUG,
                        MessageCode := 0,
                        MessageText := 'Create command payload with {1} parameter(s) :',
                        Para1       := DINT_TO_STRING(ParameterCnt));
  

// Return if no parameter is remaining...
IF ( ParameterCnt = 0 ) THEN RETURN; END_IF
// dec remaining parameter(s)                        
ParameterCnt := ParameterCnt - 1;
// Create log entry for ToolNo
CreateLogMessagePara1 ( Timestamp   := AxesGroup.State.SystemTime,
                        MessageType := MessageType.CMD,
                        Severity    := Severity.DEBUG,
                        MessageCode := 0,
                        MessageText := 'Command.ToolNo = {1}',
                        Para1       :=  INT_TO_STRING(_command.ToolNo));
END_METHOD

METHOD FB_init : BOOL
VAR_INPUT
  /// if TRUE, the retain variables are initialized (warm start / cold start)
  bInitRetains : BOOL; 
  /// if TRUE, the instance afterwards gets moved into the copy code (online change)
  bInCopyCode  : BOOL;  
END_VAR
MyType := 'MC_ReadToolDataFB';

ExecMode := ExecutionMode.PARALLEL;
Priority := PriorityLevel.NORMAL;
END_METHOD

METHOD PROTECTED OnApplyOutCmd
VAR_INPUT
  /// Command message state
  State : CmdMessageState;
END_VAR
IF ( State = CmdMessageState.EMPTY ) 
THEN
  // Reset command outputs
  SysDepMemSet(pDest := ADR(OutCmd), Value := 0, DataLen := SIZEOF(OutCmd));         
END_IF

IF (( State = CmdMessageState.ACTIVE ) OR
    ( State = CmdMessageState.DONE   ))
THEN
  // Update results
  OutCmd.ToolData     := _response.ToolData;
  OutCmd.ToolNoReturn := _response.ToolNoReturn;
END_IF
END_METHOD

METHOD PROTECTED OnExecRun : DINT
VAR_IN_OUT
  /// Robot assignment of function
  AxesGroup : AxesGroup; 
END_VAR

                  // call base implementation
SUPER^.OnExecRun(AxesGroup := AxesGroup);

CASE _stepCmd OF
  
  00:  IF ( _execute_R.Q ) AND ( NOT Error)  
       THEN
         // Check function is supported and parameter are valid ?
         IF (( CheckFunctionSupported( AxesGroup := AxesGroup )) AND
             ( CheckParameterValid   ( AxesGroup := AxesGroup )))
         THEN      
           // set busy flag
           Busy := TRUE;
           // Reset command outputs
           SysDepMemSet(pDest := ADR(OutCmd), Value := 0, DataLen := SIZEOF(OutCmd));         
           // apply command parameter
          _parCmd := ParCmd;
           // init parameter sequence
          _command.ParSeq := 1;
           // create command data
           CommandData := CreateCommandPayload(AxesGroup := AxesGroup);
           // Add command to active command register
          _uniqueID := AxesGroup.Acyclic.ActiveCommandRegister.AddCmd( pCommandFB := ADR(THIS^ ));     
           // set timeout
           SetTimeout(PT := _timeoutCmd, rTimer := _timerCmd);
           // inc step counter
          _stepCmd := _stepCmd + 1;
         END_IF 
       END_IF
     

  01:  // Wait for responce received
       IF ( _responseReceived )
       THEN
         // reset response received flag
        _responseReceived := FALSE;
         // update state flags
         OnUpdateStateFlags(_response.State);
         // update state flags
         OnApplyOutCmd(_response.State);

         // Done, Aborted or Error ?
         IF (_response.State >= CmdMessageState.DONE )
         THEN           
           // Update the ToolData in user defined system datas 
           IF UpdateSystemData AND ( _response.State = CmdMessageState.DONE ) // ST-FIX F16
THEN
AxesGroup.SystemData.UpdateToolData( Caller     := THIS^,
                                                SystemTime := AxesGroup.State.SystemTime,
                                                ToolNo     := OutCmd.ToolNoReturn, 
                                                ToolData   := OutCmd.ToolData);
END_IF                     
           // set timeout
           SetTimeout(PT := _timeoutCmd, rTimer := _timerCmd);
           // inc step counter
          _stepCmd := _stepCmd + 1; 
         END_IF
       END_IF


  02: IF ( NOT Execute)
      THEN
        Reset(); 
      END_IF     

ELSE
  // invalid step
  SetError( ErrorID := RobotLibraryErrorIdEnum.ERR_INVALID_STEP, Overwrite := TRUE );
END_CASE


// Reset FB
IF ( NOT Execute )
THEN
  Reset();
END_IF
END_METHOD

METHOD PROTECTED OnUpdateStateFlags
VAR_INPUT
  /// Command message state
  State : CmdMessageState;
END_VAR
// Reset State flags
Done := FALSE;

CASE State OF

  // No operation or process is active
  CmdMessageState.EMPTY               :;
  // Created but not yet started
  CmdMessageState.CREATED             :;
  // Buffered and awaiting execution
  CmdMessageState.BUFFERED            : CommandBuffered    := TRUE;
  // Buffered in planner for future execution
  CmdMessageState.BUFFERED_IN_PLANNER : CommandBuffered    := TRUE;
  // Currently active and in progress
  CmdMessageState.ACTIVE              :;                                   
  // Interrupted and awaiting continuation
  CmdMessageState.INTERRUPTED         :;    
  // Requested for abort
  CmdMessageState.ABORT_REQUEST       :;
  // Successfully completed
  CmdMessageState.DONE                : Done               := TRUE; 
                                        Busy               := FALSE;
  // Aborted before completion
  CmdMessageState.ABORTED             : Busy               := FALSE;
  // Encountered an error during execution
  CmdMessageState.ERROR               : Error              := TRUE;
                                        Busy               := FALSE;
END_CASE
END_METHOD

METHOD INTERNAL ParseResponsePayload : DINT
VAR_INPUT
  /// Response data
  ResponseData : RobotLibraryResponseDataFB;
  /// Timestamp
  Timestamp    : SystemTime;  
END_VAR
VAR
  /// Parameter count
 _parameterCnt : DINT;
END_VAR
// Table 6-190: Received CMD payload (RC to PLC) of "ReadToolData"
// --------------------------
// Header
// --------------------------
// Byte 00 : USINT   - ParSeq | State     
// Byte 01 : SINT    - AlarmMessageSeverity    
// Byte 02 : UINT    - AlarmMessageCode HB
// Byte 03 :         - AlarmMessageCode LB
// --------------------------
// Datablock
// --------------------------
// Byte 04 : IEC_DATE   ToolData.Date HW HB;
// Byte 05 :            ToolData.Date HW LB;
// Byte 06 : IEC_TIME - ToolData.Time HW HB;
// Byte 07 :            ToolData.Time HW LB;
// Byte 08 :            ToolData.Time LW HB;
// Byte 09 :            ToolData.Time LW LB;
// Byte 10 : REAL       ToolData.X HW HB;
// Byte 11 :            ToolData.X HW LB;
// Byte 12 :            ToolData.X LW HB;
// Byte 13 :            ToolData.X LW LB;
// Byte 14 : REAL       ToolData.Y HW HB;
// Byte 15 :            ToolData.Y HW LB;
// Byte 16 :            ToolData.Y LW HB;
// Byte 17 :            ToolData.Y LW LB;
// Byte 18 : REAL       ToolData.Z HW HB;
// Byte 19 :            ToolData.Z HW LB;
// Byte 20 :            ToolData.Z LW HB;
// Byte 21 :            ToolData.Z LW LB;
// Byte 22 : REAL       ToolData.RX HW HB;
// Byte 23 :            ToolData.RX HW LB;
// Byte 24 :            ToolData.RX LW HB;
// Byte 25 :            ToolData.RX LW LB;
// Byte 26 : REAL       ToolData.RY HW HB;
// Byte 27 :            ToolData.RY HW LB;
// Byte 28 :            ToolData.RY LW HB;
// Byte 29 :            ToolData.RY LW LB;
// Byte 30 : REAL       ToolData.RZ HW HB;
// Byte 31 :            ToolData.RZ HW LB;
// Byte 32 :            ToolData.RZ LW HB;
// Byte 33 :            ToolData.RZ LW LB;
// Byte 34 : USINT      ToolData.ID;
// Byte 35 : USINT      ToolData.LoadNo;
// Byte 36 : BOOL       ToolData.ExternalTCP;
// Byte 37 : BYTE       Reserved;

// order as table 6-190 of spec V1.5.9 (ST-FIX F27)
// Byte 38 : USINT      ToolNo;
// Byte 39 : BOOL       DataChanged;
// --------------------------
// call base implementation to parse the header from payload buffer
ResponseData.PayloadPtr := SUPER^.ParseResponsePayload(ResponseData := ResponseData, Timestamp := Timestamp);

// ST-FIX F100: missing (trailing zero) bytes of the payload are 0, no values of the previous response
SysDepMemSet( pDest := ADR(_response), Value := 0, DataLen := SIZEOF(_response));

// copy parsed header to response
_response.ParSeq               := _rspHeader.ParSeq;
_response.State                := _rspHeader.State;
_response.AlarmMessageSeverity := _rspHeader.AlarmMessageSeverity;
_response.AlarmMessageCode     := _rspHeader.AlarmMessageCode;


// Check payload remaining ? 
IF ( ResponseData.IsPayloadRemaining)
THEN  
  // Get Response.ToolData.Timestamp.IEC_DATE
 _response.ToolData.Timestamp.IEC_DATE := ResponseData.GetIecDate();
  // inc parameter counter
 _parameterCnt := _parameterCnt + 1;
END_IF


// Check payload remaining ? 
IF ( ResponseData.IsPayloadRemaining)
THEN  
  // Get Response.ToolData.Timestamp.IEC_TIME
 _response.ToolData.Timestamp.IEC_TIME := ResponseData.GetIecTime();
  // inc parameter counter
 _parameterCnt := _parameterCnt + 1;
END_IF


// Check payload remaining ? 
IF ( ResponseData.IsPayloadRemaining)
THEN  
  // Get Response.ToolData.X
 _response.ToolData.X := ResponseData.GetReal();
  // inc parameter counter
 _parameterCnt := _parameterCnt + 1;
END_IF


// Check payload remaining ? 
IF ( ResponseData.IsPayloadRemaining)
THEN  
  // Get Response.ToolData.Y
 _response.ToolData.Y := ResponseData.GetReal();
  // inc parameter counter
 _parameterCnt := _parameterCnt + 1;
END_IF


// Check payload remaining ? 
IF ( ResponseData.IsPayloadRemaining)
THEN  
  // Get Response.ToolData.Z
 _response.ToolData.Z := ResponseData.GetReal();
  // inc parameter counter
 _parameterCnt := _parameterCnt + 1;
END_IF


// Check payload remaining ? 
IF ( ResponseData.IsPayloadRemaining)
THEN  
  // Get Response.ToolData.Rx
 _response.ToolData.Rx := ResponseData.GetReal();
  // inc parameter counter
 _parameterCnt := _parameterCnt + 1;
END_IF


// Check payload remaining ? 
IF ( ResponseData.IsPayloadRemaining)
THEN  
  // Get Response.ToolData.Ry
 _response.ToolData.Ry := ResponseData.GetReal();
  // inc parameter counter
 _parameterCnt := _parameterCnt + 1;
END_IF


// Check payload remaining ? 
IF ( ResponseData.IsPayloadRemaining)
THEN  
  // Get Response.ToolData.Rz
 _response.ToolData.Rz := ResponseData.GetReal();
  // inc parameter counter
 _parameterCnt := _parameterCnt + 1;
END_IF


// Check payload remaining ? 
IF ( ResponseData.IsPayloadRemaining)
THEN  
  // Get Response.ToolData.ID
 _response.ToolData.ID := ResponseData.GetUsint();
  // inc parameter counter
 _parameterCnt := _parameterCnt + 1;
END_IF


// Check payload remaining ? 
IF ( ResponseData.IsPayloadRemaining)
THEN  
  // Get Response.ToolData.LoadNo
 _response.ToolData.LoadNo := ResponseData.GetUsint();
  // inc parameter counter
 _parameterCnt := _parameterCnt + 1;
END_IF


// Check payload remaining ? 
IF ( ResponseData.IsPayloadRemaining)
THEN  
  // Get Response.ToolData.ExternalTCP
 _response.ToolData.ExternalTCP := ResponseData.GetBool();
  // inc parameter counter
 _parameterCnt := _parameterCnt + 1;
END_IF


// Check payload remaining ? 
IF ( ResponseData.IsPayloadRemaining)
THEN  
  // Get Response.Reserve
 _response.Reserve := ResponseData.GetByte();
  // inc parameter counter
 _parameterCnt := _parameterCnt + 1;
END_IF

 
// ST-FIX F27: ToolNo first, then DataChanged (table 6-190 of spec V1.5.9)
// Check payload remaining ? 
IF ( ResponseData.IsPayloadRemaining)
THEN  
  // Get Response.ToolData.ToolNoReturn (ST-FIX F27)
 _response.ToolNoReturn := ResponseData.GetUsint();
  // inc parameter counter
 _parameterCnt := _parameterCnt + 1;
END_IF


// Check payload remaining ? 
IF ( ResponseData.IsPayloadRemaining)
THEN  
  // Get Response.DataChanged (ST-FIX F27)
 _response.DataChanged := ResponseData.GetBool();
  // inc parameter counter
 _parameterCnt := _parameterCnt + 1;
END_IF


// Create logging
ParseResponsePayloadLog(ResponseData := ResponseData, Timestamp := Timestamp, ParameterCnt := _parameterCnt);
END_METHOD

METHOD INTERNAL ParseResponsePayloadLog
VAR_INPUT
  /// Response data
  ResponseData : RobotLibraryResponseDataFB;
  /// Timestamp
  Timestamp    : SystemTime;  
  /// Parameter count
  ParameterCnt : DINT;
END_VAR
// Create log entry for Parameter start
CreateLogMessagePara1 ( Timestamp   := Timestamp,
                        MessageType := MessageType.CMD,
                        Severity    := Severity.DEBUG,
                        MessageCode := 0,
                        MessageText := '{1} parameter(s) to parse from the response data:',
                        Para1       := DINT_TO_STRING(ParameterCnt));                       


// Return if no parameter is remaining...
IF ( ParameterCnt = 0 ) THEN RETURN; END_IF
// dec remaining parameter(s)                        
ParameterCnt := ParameterCnt - 1;
// Create log entry for ToolData.Timestamp.IEC_DATE
CreateLogMessagePara1 ( Timestamp   := Timestamp,
                        MessageType := MessageType.CMD,
                        Severity    := Severity.DEBUG,
                        MessageCode := 0,
                        MessageText := 'Response.ToolData.Timestamp.IEC_DATE = {1}',
                        Para1       :=  IEC_DATE_TO_STRING(_response.ToolData.Timestamp.IEC_DATE));


// Return if no parameter is remaining...
IF ( ParameterCnt = 0 ) THEN RETURN; END_IF
// dec remaining parameter(s)                        
ParameterCnt := ParameterCnt - 1;
// Create log entry for ToolData.Timestamp.IEC_TIME
CreateLogMessagePara1 ( Timestamp   := Timestamp,
                        MessageType := MessageType.CMD,
                        Severity    := Severity.DEBUG,
                        MessageCode := 0,
                        MessageText := 'Response.ToolData.Timestamp.IEC_TIME = {1}',
                        Para1       :=  IEC_TIME_TO_STRING(_response.ToolData.Timestamp.IEC_TIME));


// Return if no parameter is remaining...
IF ( ParameterCnt = 0 ) THEN RETURN; END_IF
// dec remaining parameter(s)                        
ParameterCnt := ParameterCnt - 1;
// Create log entry for ToolData.X
CreateLogMessagePara1 ( Timestamp   := Timestamp,
                        MessageType := MessageType.CMD,
                        Severity    := Severity.DEBUG,
                        MessageCode := 0,
                        MessageText := 'Response.ToolData.X = {1}',
                        Para1       :=  REAL_TO_STRING(_response.ToolData.X));


// Return if no parameter is remaining...
IF ( ParameterCnt = 0 ) THEN RETURN; END_IF
// dec remaining parameter(s)                        
ParameterCnt := ParameterCnt - 1;
// Create log entry for ToolData.Y
CreateLogMessagePara1 ( Timestamp   := Timestamp,
                        MessageType := MessageType.CMD,
                        Severity    := Severity.DEBUG,
                        MessageCode := 0,
                        MessageText := 'Response.ToolData.Y = {1}',
                        Para1       :=  REAL_TO_STRING(_response.ToolData.Y));


// Return if no parameter is remaining...
IF ( ParameterCnt = 0 ) THEN RETURN; END_IF
// dec remaining parameter(s)                        
ParameterCnt := ParameterCnt - 1;
// Create log entry for ToolData.Z
CreateLogMessagePara1 ( Timestamp   := Timestamp,
                        MessageType := MessageType.CMD,
                        Severity    := Severity.DEBUG,
                        MessageCode := 0,
                        MessageText := 'Response.ToolData.Z = {1}',
                        Para1       :=  REAL_TO_STRING(_response.ToolData.Z));


// Return if no parameter is remaining...
IF ( ParameterCnt = 0 ) THEN RETURN; END_IF
// dec remaining parameter(s)                        
ParameterCnt := ParameterCnt - 1;
// Create log entry for ToolData.Rx
CreateLogMessagePara1 ( Timestamp   := Timestamp,
                        MessageType := MessageType.CMD,
                        Severity    := Severity.DEBUG,
                        MessageCode := 0,
                        MessageText := 'Response.ToolData.Rx = {1}',
                        Para1       :=  REAL_TO_STRING(_response.ToolData.Rx));


// Return if no parameter is remaining...
IF ( ParameterCnt = 0 ) THEN RETURN; END_IF
// dec remaining parameter(s)                        
ParameterCnt := ParameterCnt - 1;
// Create log entry for ToolData.Ry
CreateLogMessagePara1 ( Timestamp   := Timestamp,
                        MessageType := MessageType.CMD,
                        Severity    := Severity.DEBUG,
                        MessageCode := 0,
                        MessageText := 'Response.ToolData.Ry = {1}',
                        Para1       :=  REAL_TO_STRING(_response.ToolData.Ry));


// Return if no parameter is remaining...
IF ( ParameterCnt = 0 ) THEN RETURN; END_IF
// dec remaining parameter(s)                        
ParameterCnt := ParameterCnt - 1;
// Create log entry for ToolData.Rz
CreateLogMessagePara1 ( Timestamp   := Timestamp,
                        MessageType := MessageType.CMD,
                        Severity    := Severity.DEBUG,
                        MessageCode := 0,
                        MessageText := 'Response.ToolData.Rz = {1}',
                        Para1       :=  REAL_TO_STRING(_response.ToolData.Rz));


// Return if no parameter is remaining...
IF ( ParameterCnt = 0 ) THEN RETURN; END_IF
// dec remaining parameter(s)                        
ParameterCnt := ParameterCnt - 1;
// Create log entry for ToolData.ID
CreateLogMessagePara1 ( Timestamp   := Timestamp,
                        MessageType := MessageType.CMD,
                        Severity    := Severity.DEBUG,
                        MessageCode := 0,
                        MessageText := 'Response.ToolData.ID = {1}',
                        Para1       :=  USINT_TO_STRING(_response.ToolData.ID));


// Return if no parameter is remaining...
IF ( ParameterCnt = 0 ) THEN RETURN; END_IF
// dec remaining parameter(s)                        
ParameterCnt := ParameterCnt - 1;
// Create log entry for ToolData.LoadNo
CreateLogMessagePara1 ( Timestamp   := Timestamp,
                        MessageType := MessageType.CMD,
                        Severity    := Severity.DEBUG,
                        MessageCode := 0,
                        MessageText := 'Response.ToolData.LoadNo = {1}',
                        Para1       :=  USINT_TO_STRING(_response.ToolData.LoadNo));


// Return if no parameter is remaining...
IF ( ParameterCnt = 0 ) THEN RETURN; END_IF
// dec remaining parameter(s)                        
ParameterCnt := ParameterCnt - 1;
// Create log entry for ToolData.ExternalTCP
CreateLogMessagePara1 ( Timestamp   := Timestamp,
                        MessageType := MessageType.CMD,
                        Severity    := Severity.DEBUG,
                        MessageCode := 0,
                        MessageText := 'Response.ToolData.ExternalTCP = {1}',
                        Para1       :=  BOOL_TO_STRING(_response.ToolData.ExternalTCP));


// Return if no parameter is remaining...
IF ( ParameterCnt = 0 ) THEN RETURN; END_IF
// dec remaining parameter(s)                        
ParameterCnt := ParameterCnt - 1;
// Create log entry for Reserve
CreateLogMessagePara1 ( Timestamp   := Timestamp,
                        MessageType := MessageType.CMD,
                        Severity    := Severity.DEBUG,
                        MessageCode := 0,
                        MessageText := 'Response.Reserve = {1}',
                        Para1       :=  BYTE_TO_STRING(_response.Reserve));


// Return if no parameter is remaining...
IF ( ParameterCnt = 0 ) THEN RETURN; END_IF
// dec remaining parameter(s)                        
ParameterCnt := ParameterCnt - 1;
// Create log entry for ToolNoReturn
CreateLogMessagePara1 ( Timestamp   := Timestamp,
                        MessageType := MessageType.CMD,
                        Severity    := Severity.DEBUG,
                        MessageCode := 0,
                        MessageText := 'Response.ToolNoReturn = {1}',
                        Para1       :=  USINT_TO_STRING(_response.ToolNoReturn));


// Return if no parameter is remaining...
IF ( ParameterCnt = 0 ) THEN RETURN; END_IF
// dec remaining parameter(s)                        
ParameterCnt := ParameterCnt - 1;
// Create log entry for DataChanged
CreateLogMessagePara1 ( Timestamp   := Timestamp,
                        MessageType := MessageType.CMD,
                        Severity    := Severity.DEBUG,
                        MessageCode := 0,
                        MessageText := 'Response.DataChanged = {1}',
                        Para1       :=  BOOL_TO_STRING(_response.DataChanged));
END_METHOD

METHOD PROTECTED Reset : DINT
VAR_INPUT
END_VAR
Reset := SUPER^.Reset();

Done               := FALSE;
Busy               := FALSE;
CommandBuffered    := FALSE;
END_METHOD

END_FUNCTION_BLOCK

// Library/POUs/Read/MC_ReadFrameData/MC_ReadFrameDataFB

            
              /// Read content of selected user frame number
FUNCTION_BLOCK MC_ReadFrameDataFB EXTENDS RobotLibraryBaseExecuteFB
// ------------------------------------------------------------------------- 
//  SRCI Robot Library                                                
// ------------------------------------------------------------------------- 
//                                                                           
//  Object:      ReadFrameDataFB                                       
//  Author:      Thorsten Brach                                                
//  Date:        2024-06-01
//
//  Description:                                              
//   
//                                                                           
//  Copyright: 
//    (C) 2024 Thorsten Brach. All rights reserved                                                                                                                                            
//             Licensed under the MIT License.
//                                                                           
//  Disclaimer:                                                                           
//    This project is provided without any guarantee and can be used for   
//    private and commercial purposes. Any use is at the user’s 
//    own risk and responsibility.
//
// -------------------------------------------------------------------------
VAR_INPUT
  /// command parameter 
  ParCmd          : ReadFrameDataParCmd;
END_VAR
VAR_OUTPUT
  /// Command is transferred and confirmed by the RC
  CommandBuffered : BOOL;
  /// command outputs
  OutCmd          : ReadFrameDataOutCmd;       
END_VAR

VAR
  /// internal copy of command parameter 
 _parCmd          : ReadFrameDataParCmd;
  /// command data to send
 _command         : ReadFrameDataSendData;
  /// response data received
 _response        : ReadFrameDataRecvData;      
END_VAR
            
          
VAR_INPUT
  UpdateSystemData : BOOL := TRUE; // ST-FIX F16: FALSE for the internal instances of MC_RobotTaskFB (synchronisation)
END_VAR

SUPER^(AxesGroup := AxesGroup);

METHOD INTERNAL CheckAddParameter : BOOL
VAR_INPUT
  /// Payload pointer
  PayloadPtr : UDINT;
END_VAR
VAR
  /// Payload as byte array
  Payload    : ARRAY [1..SIZEOF(_command)] OF BYTE;
  /// Null Byte array 
  Null       : ARRAY [1..SIZEOF(_command)] OF BYTE;
  /// Data length to compare
  DataLen    : UDINT;
END_VAR
// Payload pointer must be decreased by one byte, because ADR(Payload) is already one byte !
PayloadPtr := LIMIT (0, PayloadPtr - 1, SIZEOF(Payload) -1);
// Convert command struct to payload array
SysDepMemCpy( pDest := ADR(Payload), pSrc := ADR(_command), DataLen := SIZEOF(_command));
// Calculate the data length to compare - at least one byte must be compared !
DataLen := LIMIT(1, SIZEOF(Payload) - PayloadPtr, SIZEOF(Payload)); 
// Compare Payload-Array with Null-Byte-Array
CheckAddParameter := SysDepMemCmp( pData1 := ADR(Payload) + PayloadPtr , pData2 := ADR(Null), DataLen := DataLen) <>  RobotLibraryConstants.OK ;
END_METHOD

METHOD PROTECTED CheckFunctionSupported : BOOL
VAR_IN_OUT
  /// Robot assignment of function
  AxesGroup : AxesGroup; 
END_VAR
CheckFunctionSupported := AxesGroup.State.RobotData.RCSupportedFunctions.ReadFrameData;

IF ( NOT CheckFunctionSupported )
THEN
  // call base implementation for set error and create log entry
  SUPER^.CheckFunctionSupported(AxesGroup := AxesGroup);
END_IF
END_METHOD

METHOD PROTECTED CheckParameterChanged : BOOL
VAR_IN_OUT
  /// Robot assignment of function
  AxesGroup    : AxesGroup; 
END_VAR
// Check ParCmd Size is > 0, because MemCmp does not work correctly with size = 0
IF (SIZEOF(ParCmd) = 0) OR (_stepCmd = 0)
THEN 
  RETURN;
END_IF

// compare memory 
_parameterChanged := ( SysDepMemCmp(pData1 := ADR(ParCmd), pData2 := ADR(_parCmd), DataLen := SIZEOF(ParCmd)) <> RobotLibraryConstants.OK );

// check parameter valid ?
_parameterValid   := CheckParameterValid( AxesGroup := AxesGroup );

IF ((  _parameterChanged        )  AND 
    (  _parameterValid          )) OR
    (  _parameterUpdateInternal )  
THEN  
  // Create log entry for parameter changed event
  CreateLogMessagePara1 ( Timestamp   := AxesGroup.State.SystemTime,
                          MessageType := MessageType.CMD,
                          Severity    := Severity.DEBUG,
                          MessageCode := 0,
                          MessageText := 'NotifyParameterChanged Event {1}',
                          Para1       :=  '' );

  // reset internal flag for send parameter update
 _parameterUpdateInternal := FALSE;
  // update internal copy of parameters 
 _parCmd := ParCmd;
  // inc parameter sequence
 _command.ParSeq := _command.ParSeq + 1;
  // update command data  
  CommandData := CreateCommandPayload(AxesGroup := AxesGroup); // ( Access via reference to rCommandFB in ACR )
  // notify active command register 
  AxesGroup.Acyclic.ActiveCommandRegister.NotifyParameterChanged := _uniqueID;
END_IF
END_METHOD

METHOD PROTECTED CheckParameterValid : BOOL
VAR_IN_OUT
  /// Robot assignment of function
  AxesGroup : AxesGroup; 
END_VAR
VAR
  /// internal index for loops
 _idx : DINT;
END_VAR
CheckParameterValid := TRUE;

// Check ParCmd.FrameNo valid ? 
IF (( ParCmd.FrameNo <  -1                                                 ) OR  
    ( ParCmd.FrameNo > 254                                                 ) OR
    ( ParCmd.FrameNo > AxesGroup.State.ConfigurationData.HighestFrameIndex ) OR
    ( ParCmd.FrameNo > AxesGroup.State.UnifiedFrameIndex                   ))         
THEN
  // Parameter not valid
  CheckParameterValid := FALSE;
  
  // Check FrameNo available on RC ? 
  IF (( ParCmd.FrameNo > AxesGroup.State.ConfigurationData.HighestFrameIndex ) AND ( ParCmd.FrameNo <= 254 )) // ST-FIX F98: outside -1..254 is a range error
  THEN
    SetError( ErrorID := RobotLibraryErrorIdEnum.ERR_FRAMENO_UNAVAILABLE, Overwrite := TRUE );
  ELSE
    SetError( ErrorID := RobotLibraryErrorIdEnum.ERR_FRAMENO_RANGE, Overwrite := TRUE );
	END_IF  
  
  // Create log entry
  CreateLogMessagePara1 ( Timestamp   := AxesGroup.State.SystemTime,
                          MessageType := MessageType.CMD,
                          Severity    := Severity.ERROR,
                          MessageCode := ErrorID,
                          MessageText := 'Invalid Parameter ParCmd.FrameNo = {1}',
                          Para1       :=  INT_TO_STRING(ParCmd.FrameNo));
  RETURN;                          
END_IF
END_METHOD

METHOD INTERNAL CreateCommandPayload : RobotLibraryCommandDataFB
VAR_IN_OUT
  /// Robot assignment of function
  AxesGroup : AxesGroup; 
END_VAR
VAR
  /// Parameter count
 _parameterCnt : DINT;
END_VAR
// Table 6-183: Sent CMD payload (PLC to RC) of "ReadFrameData"
// --------------------------
// Header
// --------------------------
// Byte 00 : UINT  - Type HB     
// Byte 01 :       - Type LB    
// Byte 02 : USINT - Reserve | ExecutionMode
// Byte 03 : USINT - ParSeq  | Priority
// --------------------------
// Datablock
// --------------------------
// Byte 04 : USINT - FrameNo
// --------------------------
// set command parameter 
_command.CmdTyp   :=  CmdType.ReadFrameData;
_command.ExecMode :=  ExecMode;
_command.ParSeq   := _command.ParSeq;
_command.Priority :=  Priority;
_command.FrameNo  :=  INT_TO_USINT(_parCmd.FrameNo);

IF (_parCmd.FrameNo = -1)
THEN
  _command.FrameNo := 255; // -1 is mapped to 255, see specification
END_IF


// copy command data to header
_cmdHeader := _command;
// call base implementation to copy header to payload buffer
CreateCommandPayload := SUPER^.CreateCommandPayload(AxesGroup := AxesGroup);


// Check parameter must be added ? 
IF ( CheckAddParameter(CreateCommandPayload.PayloadPtr))
THEN
  // add command.FrameNo
  CreateCommandPayload.AddUsint(_command.FrameNo);
  // inc parameter counter
 _parameterCnt := _parameterCnt + 1;  
END_IF


// Create logging
CreateCommandPayloadLog(AxesGroup := AxesGroup, ParameterCnt := _parameterCnt);
END_METHOD

METHOD INTERNAL CreateCommandPayloadLog
VAR_IN_OUT
  /// Robot assignment of function
  AxesGroup : AxesGroup; 
END_VAR
VAR_INPUT
  /// Parameter count
  ParameterCnt : DINT;
END_VAR
// Create log entry for Parameter start
CreateLogMessagePara1 ( Timestamp   := AxesGroup.State.SystemTime,
                        MessageType := MessageType.CMD,
                        Severity    := Severity.DEBUG,
                        MessageCode := 0,
                        MessageText := 'Create command payload with {1} parameter(s) :',
                        Para1       := DINT_TO_STRING(ParameterCnt));
  

// Return if no parameter is remaining...
IF ( ParameterCnt = 0 ) THEN RETURN; END_IF
// dec remaining parameter(s)                        
ParameterCnt := ParameterCnt - 1;
// Create log entry for FrameNo
CreateLogMessagePara1 ( Timestamp   := AxesGroup.State.SystemTime,
                        MessageType := MessageType.CMD,
                        Severity    := Severity.DEBUG,
                        MessageCode := 0,
                        MessageText := 'Command.FrameNo = {1}',
                        Para1       :=  INT_TO_STRING(_command.FrameNo));
END_METHOD

METHOD FB_init : BOOL
VAR_INPUT
  /// if TRUE, the retain variables are initialized (warm start / cold start)
  bInitRetains : BOOL; 
  /// if TRUE, the instance afterwards gets moved into the copy code (online change)
  bInCopyCode  : BOOL;  
END_VAR
MyType := 'MC_ReadFrameDataFB';

ExecMode := ExecutionMode.PARALLEL;
Priority := PriorityLevel.NORMAL;
END_METHOD

METHOD PROTECTED OnApplyOutCmd
VAR_INPUT
  /// Command message state
  State : CmdMessageState;
END_VAR
IF ( State = CmdMessageState.EMPTY ) 
THEN
  // Reset command outputs
  SysDepMemSet(pDest := ADR(OutCmd), Value := 0, DataLen := SIZEOF(OutCmd));         
END_IF

IF (( State = CmdMessageState.ACTIVE ) OR
    ( State = CmdMessageState.DONE   ))
THEN
  // Update results
  OutCmd.FrameData     := _response.FrameData;
  OutCmd.FrameNoReturn := _response.FrameNoReturn;
END_IF
END_METHOD

METHOD PROTECTED OnExecRun : DINT
VAR_IN_OUT
  /// Robot assignment of function
  AxesGroup : AxesGroup; 
END_VAR

                  // call base implementation
SUPER^.OnExecRun(AxesGroup := AxesGroup);

CASE _stepCmd OF
  
  00:  IF ( _execute_R.Q ) AND ( NOT Error)  
       THEN
         // Check function is supported and parameter are valid ?
         IF (( CheckFunctionSupported( AxesGroup := AxesGroup )) AND
             ( CheckParameterValid   ( AxesGroup := AxesGroup )))
         THEN      
           // set busy flag
           Busy := TRUE;
           // Reset command outputs
           SysDepMemSet(pDest := ADR(OutCmd), Value := 0, DataLen := SIZEOF(OutCmd));         
           // apply command parameter
          _parCmd := ParCmd;
           // init parameter sequence
          _command.ParSeq := 1;
           // create command data
           CommandData := CreateCommandPayload(AxesGroup := AxesGroup);
           // Add command to active command register
          _uniqueID := AxesGroup.Acyclic.ActiveCommandRegister.AddCmd( pCommandFB := ADR(THIS^ ));     
           // set timeout
           SetTimeout(PT := _timeoutCmd, rTimer := _timerCmd);
           // inc step counter
          _stepCmd := _stepCmd + 1;
         END_IF 
       END_IF
     

  01:  // Wait for responce received
       IF ( _responseReceived )
       THEN
         // reset response received flag
        _responseReceived := FALSE;
         // update state flags
         OnUpdateStateFlags(_response.State);
         // update state flags
         OnApplyOutCmd(_response.State);
                
         // Done, Aborted or Error ?
         IF (_response.State >= CmdMessageState.DONE )
         THEN
           // Update the FrameData in user defined system data 
           IF UpdateSystemData AND ( _response.State = CmdMessageState.DONE ) // ST-FIX F16
THEN
AxesGroup.SystemData.UpdateFrameData( Caller     := THIS^,
                                                 SystemTime := AxesGroup.State.SystemTime,
                                                 FrameNo    := OutCmd.FrameNoReturn, 
                                                 FrameData  := OutCmd.FrameData);
END_IF
           // set timeout
           SetTimeout(PT := _timeoutCmd, rTimer := _timerCmd);
           // inc step counter
          _stepCmd := _stepCmd + 1; 
         END_IF
       END_IF


  02: IF ( NOT Execute)
      THEN
        Reset();
      END_IF     

ELSE
  // invalid step
  SetError( ErrorID := RobotLibraryErrorIdEnum.ERR_INVALID_STEP, Overwrite := TRUE );
END_CASE


// Reset FB
IF ( NOT Execute )
THEN
  Reset(); 
END_IF
END_METHOD

METHOD PROTECTED OnUpdateStateFlags
VAR_INPUT
  /// Command message state
  State : CmdMessageState;
END_VAR
// Reset State flags
Done := FALSE;

CASE State OF

  // No operation or process is active
  CmdMessageState.EMPTY               :;
  // Created but not yet started
  CmdMessageState.CREATED             :;
  // Buffered and awaiting execution
  CmdMessageState.BUFFERED            : CommandBuffered    := TRUE;
  // Buffered in planner for future execution
  CmdMessageState.BUFFERED_IN_PLANNER : CommandBuffered    := TRUE;
  // Currently active and in progress
  CmdMessageState.ACTIVE              :;                                       
  // Interrupted and awaiting continuation
  CmdMessageState.INTERRUPTED         :; 
  // Requested for abort
  CmdMessageState.ABORT_REQUEST       :;
  // Successfully completed
  CmdMessageState.DONE                : Done               := TRUE;
                                        Busy               := FALSE;
  // Aborted before completion
  CmdMessageState.ABORTED             : Busy               := FALSE;
  // Encountered an error during execution
  CmdMessageState.ERROR               : Error              := TRUE;
                                        Busy               := FALSE;
END_CASE
END_METHOD

METHOD INTERNAL ParseResponsePayload : DINT
VAR_INPUT
  /// Response data
  ResponseData : RobotLibraryResponseDataFB;
  /// Timestamp
  Timestamp    : SystemTime;  
END_VAR
VAR
  /// Parameter count
 _parameterCnt : DINT;
END_VAR
// Table 6-501: Received CMD payload (RC to PLC) of "ReadDigitalInputs"
// --------------------------
// Header
// --------------------------
// Byte 00 : USINT   - ParSeq | State     
// Byte 01 : SINT    - AlarmMessageSeverity    
// Byte 02 : UINT    - AlarmMessageCode HB
// Byte 03 :         - AlarmMessageCode LB
// --------------------------
// Datablock
// --------------------------
// Byte 04 : DATE    - FrameData.Date HW HB;
// Byte 05 :         - FrameData.Date HW LB;
// Byte 06 : TOD     - FrameData.Time HW HB;
// Byte 07 :         - FrameData.Time HW LB;
// Byte 08 :         - FrameData.Time LW HB;
// Byte 09 :         - FrameData.Time LW LB;
// Byte 10 : USINT   - FrameData.ReferenceFrame;
// Byte 11 : BYTE    - Reserved;
// Byte 12 : REAL    - FrameData.X HW HB;
// Byte 13 :         - FrameData.X HW LB;
// Byte 14 :         - FrameData.X LW HB;
// Byte 15 :         - FrameData.X LW LB;
// Byte 16 : REAL    - FrameData.Y HW HB;
// Byte 17 :         - FrameData.Y HW LB;
// Byte 18 :         - FrameData.Y LW HB;
// Byte 19 :         - FrameData.Y LW LB;
// Byte 20 : REAL    - FrameData.Z HW HB;
// Byte 21 :         - FrameData.Z HW LB;
// Byte 22 :         - FrameData.Z LW HB;
// Byte 23 :         - FrameData.Z LW LB;
// Byte 24 : REAL    - FrameData.RX HW HB;
// Byte 25 :         - FrameData.RX HW LB;
// Byte 26 :         - FrameData.RX LW HB;
// Byte 27 :         - FrameData.RX LW LB;
// Byte 28 : REAL    - FrameData.RY HW HB;
// Byte 29 :         - FrameData.RY HW LB;
// Byte 30 :         - FrameData.RY LW HB;
// Byte 31 :         - FrameData.RY LW LB;
// Byte 32 : REAL    - FrameData.RZ HW HB;
// Byte 33 :         - FrameData.RZ HW LB;
// Byte 34 :         - FrameData.RZ LW HB;
// Byte 35 :         - FrameData.RZ LW LB;
// order as table 6-184 of spec V1.5.9 (ST-FIX F27)
// Byte 36 : USINT   - FrameNo;
// Byte 37 : BOOL    - DataChanged;
// call base implementation to parse the header from payload buffer
ResponseData.PayloadPtr := SUPER^.ParseResponsePayload(ResponseData := ResponseData, Timestamp := Timestamp);

// ST-FIX F100: missing (trailing zero) bytes of the payload are 0, no values of the previous response
SysDepMemSet( pDest := ADR(_response), Value := 0, DataLen := SIZEOF(_response));

// copy parsed header to response
_response.ParSeq               := _rspHeader.ParSeq;
_response.State                := _rspHeader.State;
_response.AlarmMessageSeverity := _rspHeader.AlarmMessageSeverity;
_response.AlarmMessageCode     := _rspHeader.AlarmMessageCode;


// Check payload remaining ? 
IF ( ResponseData.IsPayloadRemaining)
THEN  
  // Get Response.FrameData.Timestamp.IEC_DATE
 _response.FrameData.Timestamp.IEC_DATE := ResponseData.GetUint();
  // inc parameter counter
 _parameterCnt := _parameterCnt + 1;
END_IF


// Check payload remaining ? 
IF ( ResponseData.IsPayloadRemaining)
THEN  
  // Get Response.FrameData.Timestamp.IEC_TIME
 _response.FrameData.Timestamp.IEC_TIME := ResponseData.GetIecTime();
  // inc parameter counter
 _parameterCnt := _parameterCnt + 1;
END_IF


// Check payload remaining ? 
IF ( ResponseData.IsPayloadRemaining)
THEN  
  // Get Response.FrameData.ReferenceFrame
_response.FrameData.ReferenceFrame := ResponseData.GetUsint();
  // inc parameter counter
 _parameterCnt := _parameterCnt + 1;
END_IF


// Check payload remaining ? 
IF ( ResponseData.IsPayloadRemaining)
THEN  
  // Get Response.FrameData.Reserve
_response.Reserve := ResponseData.GetByte();
  // inc parameter counter
 _parameterCnt := _parameterCnt + 1;
END_IF


// Check payload remaining ? 
IF ( ResponseData.IsPayloadRemaining)
THEN  
  // Get Response.FrameData.X
 _response.FrameData.X := ResponseData.GetReal();
  // inc parameter counter
 _parameterCnt := _parameterCnt + 1;
END_IF


// Check payload remaining ? 
IF ( ResponseData.IsPayloadRemaining)
THEN  
  // Get Response.FrameData.Y
 _response.FrameData.Y := ResponseData.GetReal();
  // inc parameter counter
 _parameterCnt := _parameterCnt + 1;
END_IF


// Check payload remaining ? 
IF ( ResponseData.IsPayloadRemaining)
THEN  
  // Get Response.FrameData.Z
 _response.FrameData.Z := ResponseData.GetReal();
  // inc parameter counter
 _parameterCnt := _parameterCnt + 1;
END_IF


// Check payload remaining ? 
IF ( ResponseData.IsPayloadRemaining)
THEN  
  // Get Response.FrameData.Rx
 _response.FrameData.Rx := ResponseData.GetReal();
  // inc parameter counter
 _parameterCnt := _parameterCnt + 1;
END_IF


// Check payload remaining ? 
IF ( ResponseData.IsPayloadRemaining)
THEN  
  // Get Response.FrameData.Ry
 _response.FrameData.Ry := ResponseData.GetReal();
  // inc parameter counter
 _parameterCnt := _parameterCnt + 1;
END_IF


// Check payload remaining ? 
IF ( ResponseData.IsPayloadRemaining)
THEN  
  // Get Response.FrameData.Rz
 _response.FrameData.Rz := ResponseData.GetReal();
  // inc parameter counter
 _parameterCnt := _parameterCnt + 1;
END_IF


// ST-FIX F27: FrameNo first, then DataChanged (table 6-184 of spec V1.5.9)

// Check payload remaining ? 
IF ( ResponseData.IsPayloadRemaining)
THEN  
  // Get Response.FrameNoReturn (ST-FIX F27)
 _response.FrameNoReturn := ResponseData.GetUsint();
  // inc parameter counter
 _parameterCnt := _parameterCnt + 1;
END_IF


// Check payload remaining ? 
IF ( ResponseData.IsPayloadRemaining)
THEN  
  // Get Response.DataChanged (ST-FIX F27)
 _response.DataChanged := ResponseData.GetBool();
  // inc parameter counter
 _parameterCnt := _parameterCnt + 1;
END_IF


// Create logging
ParseResponsePayloadLog(ResponseData := ResponseData, Timestamp := Timestamp, ParameterCnt := _parameterCnt);
END_METHOD

METHOD INTERNAL ParseResponsePayloadLog
VAR_INPUT
  /// Response data
  ResponseData : RobotLibraryResponseDataFB;
  /// Timestamp
  Timestamp    : SystemTime;  
  /// Parameter count
  ParameterCnt : DINT;
END_VAR
// Create log entry for Parameter start
CreateLogMessagePara1 ( Timestamp   := Timestamp,
                        MessageType := MessageType.CMD,
                        Severity    := Severity.DEBUG,
                        MessageCode := 0,
                        MessageText := '{1} parameter(s) to parse from the response data:',
                        Para1       := DINT_TO_STRING(ParameterCnt));
                        

// Return if no parameter is remaining...
IF ( ParameterCnt = 0 ) THEN RETURN; END_IF
// dec remaining parameter(s)                        
ParameterCnt := ParameterCnt - 1;
// Create log entry for FrameData.Timestamp.IEC_DATE
CreateLogMessagePara1 ( Timestamp   := Timestamp,
                        MessageType := MessageType.CMD,
                        Severity    := Severity.DEBUG,
                        MessageCode := 0,
                        MessageText := 'Response.FrameData.Timestamp.IEC_DATE = {1}',
                        Para1       :=  IEC_DATE_TO_STRING(_response.FrameData.Timestamp.IEC_DATE));


// Return if no parameter is remaining...
IF ( ParameterCnt = 0 ) THEN RETURN; END_IF
// dec remaining parameter(s)                        
ParameterCnt := ParameterCnt - 1;
// Create log entry for FrameData.Timestamp.IEC_TIME
CreateLogMessagePara1 ( Timestamp   := Timestamp,
                        MessageType := MessageType.CMD,
                        Severity    := Severity.DEBUG,
                        MessageCode := 0,
                        MessageText := 'Response.FrameData.Timestamp.IEC_TIME = {1}',
                        Para1       :=  IEC_TIME_TO_STRING(_response.FrameData.Timestamp.IEC_TIME));


// Return if no parameter is remaining...
IF ( ParameterCnt = 0 ) THEN RETURN; END_IF
// dec remaining parameter(s)                        
ParameterCnt := ParameterCnt - 1;
// Create log entry for FrameData.ReferenceFrame
CreateLogMessagePara1 ( Timestamp   := Timestamp,
                        MessageType := MessageType.CMD,
                        Severity    := Severity.DEBUG,
                        MessageCode := 0,
                        MessageText := 'Response.FrameData.ReferenceFrame = {1}',
                        Para1       :=  USINT_TO_STRING(_response.FrameData.ReferenceFrame));


// Return if no parameter is remaining...
IF ( ParameterCnt = 0 ) THEN RETURN; END_IF
// dec remaining parameter(s)                        
ParameterCnt := ParameterCnt - 1;
// Create log entry for Reserve
CreateLogMessagePara1 ( Timestamp   := Timestamp,
                        MessageType := MessageType.CMD,
                        Severity    := Severity.DEBUG,
                        MessageCode := 0,
                        MessageText := 'Response.Reserve = {1}',
                        Para1       :=  USINT_TO_STRING(_response.Reserve));


// Return if no parameter is remaining...
IF ( ParameterCnt = 0 ) THEN RETURN; END_IF
// dec remaining parameter(s)                        
ParameterCnt := ParameterCnt - 1;
// Create log entry for FrameData.X
CreateLogMessagePara1 ( Timestamp   := Timestamp,
                        MessageType := MessageType.CMD,
                        Severity    := Severity.DEBUG,
                        MessageCode := 0,
                        MessageText := 'Response.FrameData.X = {1}',
                        Para1       :=  REAL_TO_STRING(_response.FrameData.X));


// Return if no parameter is remaining...
IF ( ParameterCnt = 0 ) THEN RETURN; END_IF
// dec remaining parameter(s)                        
ParameterCnt := ParameterCnt - 1;
// Create log entry for FrameData.Y
CreateLogMessagePara1 ( Timestamp   := Timestamp,
                        MessageType := MessageType.CMD,
                        Severity    := Severity.DEBUG,
                        MessageCode := 0,
                        MessageText := 'Response.FrameData.Y = {1}',
                        Para1       :=  REAL_TO_STRING(_response.FrameData.Y));


// Return if no parameter is remaining...
IF ( ParameterCnt = 0 ) THEN RETURN; END_IF
// dec remaining parameter(s)                        
ParameterCnt := ParameterCnt - 1;
// Create log entry for FrameData.Z
CreateLogMessagePara1 ( Timestamp   := Timestamp,
                        MessageType := MessageType.CMD,
                        Severity    := Severity.DEBUG,
                        MessageCode := 0,
                        MessageText := 'Response.FrameData.Z = {1}',
                        Para1       :=  REAL_TO_STRING(_response.FrameData.Z));


// Return if no parameter is remaining...
IF ( ParameterCnt = 0 ) THEN RETURN; END_IF
// dec remaining parameter(s)                        
ParameterCnt := ParameterCnt - 1;
// Create log entry for FrameData.Rx
CreateLogMessagePara1 ( Timestamp   := Timestamp,
                        MessageType := MessageType.CMD,
                        Severity    := Severity.DEBUG,
                        MessageCode := 0,
                        MessageText := 'Response.FrameData.Rx = {1}',
                        Para1       :=  REAL_TO_STRING(_response.FrameData.Rx));


// Return if no parameter is remaining...
IF ( ParameterCnt = 0 ) THEN RETURN; END_IF
// dec remaining parameter(s)                        
ParameterCnt := ParameterCnt - 1;
// Create log entry for FrameData.Ry
CreateLogMessagePara1 ( Timestamp   := Timestamp,
                        MessageType := MessageType.CMD,
                        Severity    := Severity.DEBUG,
                        MessageCode := 0,
                        MessageText := 'Response.FrameData.Ry = {1}',
                        Para1       :=  REAL_TO_STRING(_response.FrameData.Ry));


// Return if no parameter is remaining...
IF ( ParameterCnt = 0 ) THEN RETURN; END_IF
// dec remaining parameter(s)                        
ParameterCnt := ParameterCnt - 1;
// Create log entry for FrameData.Rz
CreateLogMessagePara1 ( Timestamp   := Timestamp,
                        MessageType := MessageType.CMD,
                        Severity    := Severity.DEBUG,
                        MessageCode := 0,
                        MessageText := 'Response.FrameData.Rz = {1}',
                        Para1       :=  REAL_TO_STRING(_response.FrameData.Rz));


// Return if no parameter is remaining...
IF ( ParameterCnt = 0 ) THEN RETURN; END_IF
// dec remaining parameter(s)                        
ParameterCnt := ParameterCnt - 1;
// Create log entry for FrameNoReturn
CreateLogMessagePara1 ( Timestamp   := Timestamp,
                        MessageType := MessageType.CMD,
                        Severity    := Severity.DEBUG,
                        MessageCode := 0,
                        MessageText := 'Response.FrameNoReturn = {1}',
                        Para1       :=  USINT_TO_STRING(_response.FrameNoReturn));


// Return if no parameter is remaining...
IF ( ParameterCnt = 0 ) THEN RETURN; END_IF
// dec remaining parameter(s)                        
ParameterCnt := ParameterCnt - 1;
// Create log entry for DataChanged
CreateLogMessagePara1 ( Timestamp   := Timestamp,
                        MessageType := MessageType.CMD,
                        Severity    := Severity.DEBUG,
                        MessageCode := 0,
                        MessageText := 'Response.DataChanged = {1}',
                        Para1       :=  BOOL_TO_STRING(_response.DataChanged));
END_METHOD

METHOD PROTECTED Reset : DINT
VAR_INPUT
END_VAR
Reset := SUPER^.Reset();

Done               := FALSE;
Busy               := FALSE;
CommandBuffered    := FALSE;
END_METHOD

END_FUNCTION_BLOCK

// Library/POUs/Read/MC_ReadLoadData/MC_ReadLoadDataFB

            
              /// Read content of selected payload number
FUNCTION_BLOCK MC_ReadLoadDataFB EXTENDS RobotLibraryBaseExecuteFB
// ------------------------------------------------------------------------- 
//  SRCI Robot Library                                                
// ------------------------------------------------------------------------- 
//                                                                           
//  Object:      ReadLoadDataFB                                       
//  Author:      Thorsten Brach                                                
//  Date:        2024-06-01
//
//  Description:                                              
//   
//                                                                           
//  Copyright: 
//    (C) 2024 Thorsten Brach. All rights reserved                                                                                                                                            
//             Licensed under the MIT License.
//                                                                           
//  Disclaimer:                                                                           
//    This project is provided without any guarantee and can be used for   
//    private and commercial purposes. Any use is at the user’s 
//    own risk and responsibility.
//
// -------------------------------------------------------------------------
VAR_INPUT
  /// command parameter 
  ParCmd          : ReadLoadDataParCmd;
END_VAR
VAR_OUTPUT
  /// Command is transferred and confirmed by the RC
  CommandBuffered : BOOL;
  /// command outputs
  OutCmd          : ReadLoadDataOutCmd;       
END_VAR

VAR
  /// internal copy of command parameter 
 _parCmd          : ReadLoadDataParCmd;
  /// command data to send
 _command         : ReadLoadDataSendData;
  /// response data received
 _response        : ReadLoadDataRecvData;      
END_VAR
            
          
VAR_INPUT
  UpdateSystemData : BOOL := TRUE; // ST-FIX F16: FALSE for the internal instances of MC_RobotTaskFB (synchronisation)
END_VAR

SUPER^(AxesGroup := AxesGroup);

